(* IEC 61131-3 sources: IRIS-Project/LASAL CONTROL SOFTWARE/LasalProject_2025_09_12/Runtime/%LASALAPPDATA%/Runtime/Library/Loader/Source/code (part 10) *)

  OS_MT_Wait(pLogin^.hMutex);
  retval := SendLogout_TCP_nocs(pComdefT, pLogin);
  OS_MT_Signal(pLogin^.hMutex);

  UnlockLoginContext(pLogin); // wg. dem LockLoginContext2 Aufruf in dieser Funktion

END_FUNCTION
#endif

//------------------------------------------------------------------------------
// ComlinkT_InstallCallback
//------------------------------------------------------------------------------
#ifdef COMLINK_TCP_CLIENT
FUNCTION ComlinkT_InstallCallback
VAR_INPUT
    pCallback : ^void;
END_VAR
VAR
    i         : UDINT;
    pLogin    : ^loginContext;
END_VAR

  IF isClientReady < 0 THEN
    DEBUGLOG0("%010d-*** ComlinkT_InstallCallback: client is not ready");
    RETURN; // zeile geloescht laut pranz mail vom 30.01.2004
  END_IF;

  DEBUGLOG1("%010d-ComlinkT_InstallCallback: pCallback=0x%08X", pCallback$UDINT);

  FOR i := 0 TO (g_max_logins - 1) DO
    pLogin := LockLoginContext(i);
    IF pLogin <> NIL THEN
      pLogin^.pCallback := pCallback;
      UnlockLoginContext(pLogin);
    END_IF;
  END_FOR;

  g_pCallback := pCallback;

END_FUNCTION
#endif

//------------------------------------------------------------------------------
// ComlinkT_StartStopRefresh_nocs
//------------------------------------------------------------------------------
#ifdef COMLINK_TCP_CLIENT
FUNCTION ComlinkT_StartStopRefresh_nocs
VAR_INPUT
    pLogin   : ^loginContext; // connection context
    count    : UINT;
    typ      : UINT;
    res      : UDINT;
END_VAR
VAR_OUTPUT
    retval    : comlinkReason;
END_VAR
VAR
    reqMsg        : msgSsRefrReq;  // request structure for command CMD_SSREFR
    timeout_ms    : UDINT;         // timeout value for send request
    fFlush        : UDINT;
    rc            : DINT;
    rc2           : comlinkReason;
END_VAR

  retval := COMLINK_ERR_GENERAL;

  rc2 := CheckClientConnection(pLogin, #pLogin^.refrSockClnt, 0);
  IF rc2 <> COMLINK_OK THEN
    retval := rc2;
    RETURN;
  END_IF;

  // prepare the request message structure
  reqMsg.count   := count;
  reqMsg.typ     := typ;

  fFlush := 1;
  IF QUERY_FREE_TXBUF(pLogin^.refrSockClnt) < (2 * SIZEOF(reqMsg)) THEN
    DEBUGLOG0("%010d-*** ComlinkT_StartStopRefresh: send buffer shortage, next send will block");
    timeout_ms := CLIENT_TIMEOUT_REQ;
  ELSE
    timeout_ms := 0;    // timeout: non-blocking
  END_IF;

  pLogin^.accelerateCellUpdates := TRUE;

  // Send the request
  rc := SendCmdMsg(#pLogin^.refrSockClnt,
                   CMD_SSREFR,
                   0,                // Type and Ack field of command (type: request, ack: no response required)
                   #reqMsg$cMessage,
                   SIZEOF(reqMsg),
                   timeout_ms,
                   1,                // use buffered send
                   fFlush            // fFlush
                  );
  IF rc <= 0 THEN
    DEBUGLOG3("%010d-*** ComlinkT_StartStopRefresh(typ %d, count %d): SendCmdMsg failed, rc=%d", TO_UDINT(typ), TO_UDINT(count), TO_UDINT(rc));
    CloseBufferedSock(#pLogin^.refrSockClnt);
    retval := COMLINK_ERR_NOCONNECTION;
  ELSE
    DEBUG_VERBOSE3("%010d-ComlinkT_StartStopRefresh: SSREFR request sent, msgLen=%d, typ=%d, count=%d", TO_UDINT(rc), TO_UDINT(typ), TO_UDINT(count));
    retval := COMLINK_OK;
  END_IF;

END_FUNCTION
#endif

//------------------------------------------------------------------------------
// ComlinkT_StartStopRefresh
//------------------------------------------------------------------------------
#ifdef COMLINK_TCP_CLIENT
FUNCTION ComlinkT_StartStopRefresh
VAR_INPUT
    pComdef  : ^comdef;
    count    : UINT;
    typ      : UINT;
    res      : UDINT;
END_VAR
VAR_OUTPUT
    retval   : comlinkReason;
END_VAR
VAR
    pLogin        : ^loginContext; // connection context
END_VAR

  IF isClientReady < 0 THEN
    DEBUGLOG0("%010d-*** ComlinkT_StartStopRefresh: client is not ready");
    TraceMsg4Client();
    retval := COMLINK_ERR_CLIENT_NOTREADY;
    RETURN;
  END_IF;
  pLogin := pComdef^$comdefT.pLogin;
  IF pLogin = NIL THEN
    retval := COMLINK_ERR_LOGIN_REQUIRED;
    RETURN;
  END_IF;

  OS_MT_Wait(pLogin^.hMutex);
  retval := ComlinkT_StartStopRefresh_nocs(pLogin, count, typ, res);
  OS_MT_Signal(pLogin^.hMutex);

END_FUNCTION
#endif

//------------------------------------------------------------------------------
// ComlinkT_CyWork_Client - cyclic work for client
//------------------------------------------------------------------------------
#ifdef COMLINK_TCP_CLIENT
FUNCTION ComlinkT_CyWork_Client
VAR
    pLogin      : ^loginContext;
    reqMsgNop   : msgNopReq;
    rc          : DINT;
#ifndef LOADER_TCP_MODERATE
    i           : UDINT;
#endif
END_VAR

  IF (isClientReady < 0) | (loginAnz = 0) THEN
    RETURN;
  END_IF;

  TRACE_ENTRY(200);

#ifndef LOADER_TCP_MODERATE
  FOR i := 0 TO (g_max_logins - 1) DO

    pLogin := LockLoginContext(i);
#else
    pLogin := LockLoginContext(TCPCltCntr);
#endif

    IF pLogin <> NIL THEN

      TRACE_ENTRY(210);

      IF (pLogin^.cmdSockClnt.sock < 0) & (pLogin^.cmdSockClnt.pndSock >= 0) THEN
        // a pending command connection exists
        rc := Connect(pLogin^.cmdSockClnt.pndSock, pLogin^.ipAddrSrvr, pLogin^.cmdPortSrvr, 0);
        IF rc >= 0 THEN
          pLogin^.cmdSockClnt.sock    := pLogin^.cmdSockClnt.pndSock;
          pLogin^.cmdSockClnt.pndSock := INVALID_SOCKET_NUM;
          DEBUGLOG1("%010d-ComlinkT_CyWork: client connected to command server (port:%d)", pLogin^.cmdPortSrvr$UDINT);
        ELSIF rc <> TCP_NOT_READY THEN
          CloseSock(#pLogin^.cmdSockClnt.pndSock);
          DEBUGLOG2("%010d-ComlinkT_CyWork: connect to command server (port:%d) failed, rc=%d", pLogin^.cmdPortSrvr$UDINT, TO_UDINT(rc));
        END_IF;
      END_IF;

      IF (pLogin^.refrSockClnt.sock < 0) & (pLogin^.refrSockClnt.pndSock >= 0) THEN
        // a pending refresh connection exists
        rc := Connect(pLogin^.refrSockClnt.pndSock, pLogin^.ipAddrSrvr, pLogin^.cmdPortSrvr + 1, 0);
        IF rc >= 0 THEN
          pLogin^.refrSockClnt.sock    := pLogin^.refrSockClnt.pndSock;
          pLogin^.refrSockClnt.pndSock := INVALID_SOCKET_NUM;
          DEBUGLOG1("%010d-ComlinkT_CyWork: client connected to refresh server (port:%d)", (pLogin^.cmdPortSrvr + 1)$UDINT);
        ELSIF rc <> TCP_NOT_READY THEN
          CloseSock(#pLogin^.refrSockClnt.pndSock);
          DEBUGLOG2("%010d-ComlinkT_CyWork: connect to refresh server (port:%d) failed, rc=%d", (pLogin^.cmdPortSrvr + 1)$UDINT, TO_UDINT(rc));
        END_IF;
      END_IF;

      IF OS_MT_WaitCond(pLogin^.hMutex) THEN
        IF CheckClientConnection(pLogin, #pLogin^.refrSockClnt, 0) <> COMLINK_OK THEN

          TRACE_ENTRY(211);
          // poll for a response of the sessioninfo request
          PndConnListener(pLogin);

        ELSE

          TRACE_ENTRY(212);
          // flush the buffer when no transfer was in the last SMALLEST_UPD_INTERVALL ms
          IF (pLogin^.refrSockClnt.bytesInTxBuf > 0) &
             ((ops.tAbsolute - pLogin^.refrSockClnt.lastSendTime) > SMALLEST_UPD_INTERVALL) THEN
            DEBUG_VERBOSE1("%010d-ComlinkT_CyWork: initiate transfer of bufferd data (%d bytes)", pLogin^.refrSockClnt.bytesInTxBuf);
            FLUSH_TXBUF(#pLogin^.refrSockClnt);
          END_IF;

          // Send data at a regular interval to get informed when the server is not alive.
          // Without sending data at a regular interval we would recognize a connection failure
          // only when the LSE kernel initiates a transfer.
          // When we know that the server does not respond, we can initiate the reconnect procedure.
          IF (ops.tAbsolute - pLogin^.refrSockClnt.lastSendTime) > HEARTBEAT_INTERVALL THEN
            DEBUG_VERBOSE0("%010d-ComlinkT_CyWork: sending heartbeat");
            SendCmdMsg(#pLogin^.refrSockClnt, CMD_NOP, 0, #reqMsgNop$cMessage, SIZEOF(reqMsgNop), 0, 1, 1);
          END_IF;

          // send data in the buffer that is marked as unsent
          SendUnsentData(#pLogin^.refrSockClnt);

          // process incoming update cell requests
          IF ((ops.tAbsolute - pLogin^.refrSockClnt.lastUpdTime) > SMALLEST_UPD_INTERVALL) | pLogin^.accelerateCellUpdates THEN
            WHILE 1 DO
              IF UpdCellListener(pLogin) = 0 THEN
                // UpdCellListener returns 0 when no message is received
                EXIT;
              ELSE
                pLogin^.accelerateCellUpdates := FALSE;
              END_IF;
            END_WHILE;
            pLogin^.refrSockClnt.lastUpdTime := ops.tAbsolute;
          END_IF;

        END_IF;
        OS_MT_Signal(pLogin^.hMutex);
      END_IF; // OS_MT_WaitCond(pLogin^.hMutex)

      TRACE_ENTRY(219);

      UnlockLoginContext(pLogin);

    END_IF;

#ifdef LOADER_TCP_MODERATE
    TCPCltCntr += 1;
    if (TCPCltCntr = g_max_logins) then
      TCPCltCntr := 0;
    end_if;
#else
  END_FOR;
#endif

  TRACE_ENTRY(299);

END_FUNCTION
#endif

//------------------------------------------------------------------------------
// Ruft das Accept für den Command Socket auf
//------------------------------------------------------------------------------
#ifdef COMLINK_TCP_SERVER
FUNCTION ComlinkT_AcceptCmdSock
VAR
    sock        : DINT;
END_VAR

  IF cmdSockSrvr >= 0 THEN
    sock := OS_TCP_USER_ACCEPT(cmdSockSrvr, 0);
    IF sock >= 0 THEN
      DEBUGLOG1("%010d-  =====  command client connected  =====  , sock=%d", sock$UDINT);
      IF sock < arraysize(usedsocks) THEN
        usedsocks[sock] := 'C';
      END_IF;
      SetSocketOptions(sock);
      IF AllocConnBlock(TYPE_CMD_CONN, sock) = NIL THEN
        CloseSock(#sock);
      END_IF;
    END_IF;
  END_IF;

END_FUNCTION
#endif

//------------------------------------------------------------------------------
// Ruft das Accept für den Refresh Socket auf
//------------------------------------------------------------------------------
#ifdef COMLINK_TCP_SERVER
FUNCTION ComlinkT_AcceptRefrSock
VAR
    sock        : DINT;
END_VAR

  IF refrSockSrvr >= 0 THEN
    sock := OS_TCP_USER_ACCEPT(refrSockSrvr, 0);
    IF sock >= 0 THEN
      DEBUGLOG1("%010d-  =====  refresh client connected  =====  , sock=%d", sock$UDINT);
      IF sock < arraysize(usedsocks) THEN
        usedsocks[sock] := 'R';
      END_IF;
      SetSocketOptions(sock);
      IF AllocConnBlock(TYPE_REFR_CONN, sock) = NIL THEN
        CloseSock(#sock);
      END_IF;
    END_IF;
  END_IF;

END_FUNCTION
#endif

//------------------------------------------------------------------------------
// Serviciert einen offenen Command Socket
//------------------------------------------------------------------------------
#ifdef COMLINK_TCP_SERVER
FUNCTION ComlinkT_ServeCmdSock
VAR_INPUT
    pCmdConn    : ^cmdConnBlock;
END_VAR
#ifdef LOADER_TCP_MODERATE
VAR
	rc : DINT;
END_VAR
#endif

    // send data in the buffer that is marked as unsent
    SendUnsentData(#pCmdConn^.bsock);

    // process incoming command requests
    #ifdef LOADER_TCP_MODERATE
    rc :=
    #endif
    CmdMsgListener(pCmdConn);

    #ifdef LOADER_TCP_MODERATE
    IF rc >= 0 THEN
      pCmdConn^.bSock.isDataAvailable := false;
    END_IF;
    #endif

END_FUNCTION
#endif

//------------------------------------------------------------------------------
// Serviciert einen offenen Refresh Socket
//------------------------------------------------------------------------------
#ifdef COMLINK_TCP_SERVER
FUNCTION ComlinkT_ServeRefrSock
VAR_INPUT
    pRefrConn   : ^refrConnBlock;
END_VAR
VAR
    i           : UDINT;
    rc : DINT;
END_VAR

    // flush the buffer when no transfer was in the last SMALLEST_UPD_INTERVALL ms
    IF (pRefrConn^.bsock.bytesInTxBuf > 0) &
       ((ops.tAbsolute - pRefrConn^.bsock.lastSendTime) > SMALLEST_UPD_INTERVALL) THEN
      DEBUG_VERBOSE1("%010d-ComlinkT_CyWork: initiate transfer of bufferd data (%d bytes)", pRefrConn^.bsock.bytesInTxBuf);
      FLUSH_TXBUF(#pRefrConn^.bsock);
    END_IF;
    // send data in the buffer that is marked as unsent
    SendUnsentData(#pRefrConn^.bsock);

    // process incoming requests (TXUPD, StartStopRefresh)
    IF pRefrConn^.bsock.lastSendTime_ms <> ops.tAbsolute |
       pRefrConn^.bsock.refrMsgListenInhibitCnt > 5 // damit der RefrMsgListener auch eine Chance hat
       THEN
      // Es wird nur ein Receive durchgeführt, wenn in diesem Durchlauf nichts
      // gesendet wurde. Das begrenzt die CPU Last.
      i := 0;
      WHILE 1 DO
        rc := RefrMsgListener(pRefrConn);
        IF rc = 0 THEN
          // RefrMsgListener returns 0 when no message is received
          EXIT;
        END_IF;
        IF rc < 0 THEN
          // pRefrConn was released
          RETURN;
        END_IF;
        i += 1;
        IF i > 500 THEN // for safety
          EXIT;
        END_IF;
      END_WHILE;
      pRefrConn^.bsock.refrMsgListenInhibitCnt := 0;
    ELSE
      pRefrConn^.bsock.refrMsgListenInhibitCnt += 1;
    END_IF;
    // scan the update list and send changes to the client
    IF pRefrConn^.bsock.fTxBufferShortage THEN
      // no update in the case ot a buffer shortage
      IF QUERY_FREE_TXBUF(pRefrConn^.bsock) > (pRefrConn^.bsock.sizeOfTxBuf / 2) THEN
        DEBUGLOG0("%010d-ComlinkT_CyWork: leaving tx buffer shortage");
        pRefrConn^.bsock.fTxBufferShortage := 0;
      END_IF;
    ELSE
      IF ((ops.tAbsolute - pRefrConn^.bsock.lastUpdTime) > SMALLEST_UPD_INTERVALL) | pRefrConn^.flushNextSends THEN
        UpdateListProcessor(pRefrConn);
        pRefrConn^.bsock.lastUpdTime := ops.tAbsolute;
        IF pRefrConn^.flushNextSends THEN
          FLUSH_TXBUF(#pRefrConn^.bsock);
          pRefrConn^.flushNextSends := FALSE;
        END_IF;
      ELSE
        prefrconn := prefrconn;
      END_IF;
    END_IF;

    if( pRefrConn^.ptr = NIL )then
      return;
    end_if;
    IF pRefrConn^.ptr^.maxIdleTime_ms > 0 THEN
      IF ops.tAbsolute - pRefrConn^.bsock.lastSendTime_ms > pRefrConn^.ptr^.maxIdleTime_ms THEN
        SendAliveMessage_TCP(pRefrConn); // der Gegenstelle mitteilen, daß man noch lebt
      END_IF;
    END_IF;

END_FUNCTION
#endif

//------------------------------------------------------------------------------
// ComlinkT_CyWork_Server - cyclic work for server
//------------------------------------------------------------------------------
#ifdef COMLINK_TCP_SERVER
FUNCTION ComlinkT_CyWork_Server
VAR
    pCmdConnOld : ^cmdConnBlock;
    pRefrConnOld: ^refrConnBlock;
END_VAR

  IF isServerReady < 0 THEN
    RETURN;
  END_IF;

  // Die Aufrufe für das Accept des Kommando- und Refreshkanals und die
  // Bedienung dieser Kanäle wird so aufgeteilt, daß bei jedem Durchlauf
  // nur ein Aufruf gemacht wird, wobei die Accepts nur jedes 50te mal
  // aufgerufen werden. Ein Verbindungsaufbau braucht nämlich nicht so oft
  // überwacht werden.
  // Der Grund für diese Aufteilung ist der hohe CPU Verbrauch eines
  // TCP/IP Calls.

  CASE tcpServerState OF
    0:
      TRACE_ENTRY(100);
      // accept incoming command connection
      ComlinkT_AcceptCmdSock();
      tcpServerState += 1;

    1:
      TRACE_ENTRY(101);
      // accept incoming refresn connection
      ComlinkT_AcceptRefrSock();
      tcpServerState += 1;

    2:
      TRACE_ENTRY(102);
      // cyclic work for refresh server
      IF s_pRefrConn = NIL THEN
        s_pRefrConn := pRefrConnRoot;
      END_IF;
      IF s_pRefrConn <> NIL THEN

        ComlinkT_ServeRefrSock(s_pRefrConn);

        // check if an error occured
        IF s_pRefrConn <> NIL THEN // s_pRefrConn kann in ComlinkT_ServeRefrSock freigegeben werden
	        IF s_pRefrConn^.bsock.sock < 0 THEN
	          pRefrConnOld := s_pRefrConn;
	          s_pRefrConn    := s_pRefrConn^.next;
            DEBUGLOG0("%010d-  =====  Error in RefrConn -> releasing connBlock  =====");
	          ReleaseConnBlock(TYPE_REFR_CONN, pRefrConnOld$^connBlock, 1);
            pRefrConnOld := NIL;
	        ELSE
	          s_pRefrConn := s_pRefrConn^.next;
	        END_IF;
        END_IF;

      END_IF;
      IF s_pRefrConn = NIL THEN
        tcpServerState += 1;
      END_IF;

    3:
      TRACE_ENTRY(103);
      // cyclic work for command server
      IF s_pCmdConn = NIL THEN
        s_pCmdConn := pCmdConnRoot;
      END_IF;
      IF s_pCmdConn <> NIL THEN

        ComlinkT_ServeCmdSock(s_pCmdConn);

        // check if an error occured
        IF s_pCmdConn <> NIL THEN // s_pCmdConn kann in ComlinkT_ServeCmdSock freigegeben werden
	        IF s_pCmdConn^.bsock.sock < 0 THEN
	          pCmdConnOld := s_pCmdConn;
	          s_pCmdConn    := s_pCmdConn^.next;
            DEBUGLOG0("%010d-  =====  Error in CmdConn -> releasing connBlock =====");
	          ReleaseConnBlock(TYPE_CMD_CONN, pCmdConnOld$^connBlock, 0);
            pCmdConnOld := NIL;
	        ELSE
	          s_pCmdConn := s_pCmdConn^.next;
	        END_IF;
        END_IF;

      END_IF;
      IF s_pCmdConn = NIL THEN
        tcpServerState += 1;
      END_IF;

  END_CASE;

  tcpAcceptState += 1;

  IF tcpServerState > 3 THEN
    // Es wird nur alle 50 Durchläufe ein Accept eingeschoben
    IF tcpAcceptState > 50 THEN
      tcpAcceptState := 0;
      tcpServerState := 0;
    ELSE
      tcpServerState := 2;
    END_IF;
  END_IF;

  TRACE_ENTRY(199);

END_FUNCTION
#endif

//------------------------------------------------------------------------------
// ComlinkT_CyWork
//------------------------------------------------------------------------------
FUNCTION ComlinkT_CyWork

  TRACE_ENTRY(10);

#ifdef COMLINK_TCP_SERVER
  ComlinkT_CyWork_Server();
#endif

  TRACE_ENTRY(11);

#ifdef COMLINK_TCP_CLIENT
  ComlinkT_CyWork_Client();
#endif

  TRACE_ENTRY(12);

END_FUNCTION

#endif //COMLINK_TCP

#ifndef COMLINK_TCP_CLIENT

//------------------------------------------------------------------------------
// ComlinkT_MissingClientCode
//------------------------------------------------------------------------------
FUNCTION ComlinkT_MissingClientCode

  IF ComlinkT_wasTraceMsgDisplayed = 0 THEN
    TRACE_ERR("Comlink/TCP client error: missing client code (COMLINK_TCP_CLIENT not defined)");
    LSLCLI_LoaderTracePrint("Comlink/TCP client error: missing client code (COMLINK_TCP_CLIENT not defined)", 12);
    ComlinkT_wasTraceMsgDisplayed := 1;
  END_IF;

END_FUNCTION

#endif // !COMLINK_TCP_CLIENT

//++comlinkt:end

////////////////////////////////////////////////////////////////////////////////
//
//  I-am-Alive Mechanismus
//
////////////////////////////////////////////////////////////////////////////////

FUNCTION SendMaxIdleTime_CAN
VAR_INPUT
  pComdefT : ^comdefT;
  remoteMaxIdleTime_ms : UDINT;
END_VAR
VAR_OUTPUT
  retVal : DINT;
END_VAR
VAR
  txinfo4006    : COMOBJSTR;
END_VAR

    txinfo4006.iLng  := 0;
    txinfo4006.iOff  := 4006;
    txinfo4006.dData := TO_DINT(remoteMaxIdleTime_ms);

    IF CanTxObj(pComdefT$^COMDEF^.pt_COM, #txinfo4006$void) <> 0 THEN
        retVal := -1;
    ELSE
        retVal := 0;
    END_IF;

END_FUNCTION
FUNCTION SendAliveMessage_CAN
VAR_INPUT
  pCom : ^COMDATA;
END_VAR
VAR_OUTPUT
  retVal : DINT;
END_VAR
VAR
  txinfo4007    : COMOBJSTR;
END_VAR

    txinfo4007.iLng  := 0;
    txinfo4007.iOff  := 4007;
    txinfo4007.dData := 0;

    IF CanTxObj(pCom, #txinfo4007$void) <> 0 THEN
        retVal := -1;
    ELSE
        retVal := 0;
    END_IF;

END_FUNCTION
//------------------------------------------------------------------------------
// SendMaxIdleTime
//
//  Schickt die maxIdleTime zur Gegenstation
//------------------------------------------------------------------------------
FUNCTION SendMaxIdleTime
VAR_INPUT
  pComdefT : ^comdefT;
  remoteMaxIdleTime_ms : UDINT;
END_VAR
VAR_OUTPUT
  retVal : DINT;
END_VAR

  CASE pComdefT^.interface  OF

  COMLINK_IFNUM_CAN1,
  COMLINK_IFNUM_CAN2,
  COMLINK_IFNUM_CAN20,
  COMLINK_IFNUM_CAN21,
  COMLINK_IFNUM_CAN22,
  COMLINK_IFNUM_CAN23,
  COMLINK_IFNUM_CAN24,
  COMLINK_IFNUM_CAN25,
  COMLINK_IFNUM_CAN26,
  COMLINK_IFNUM_CAN27,
  COMLINK_IFNUM_CAN28,
  COMLINK_IFNUM_CAN29:
    retVal := SendMaxIdleTime_CAN(pComdefT, remoteMaxIdleTime_ms);
#ifdef COMLINK_TCP_SERVER
  COMLINK_IFNUM_TCP1_OLD,
  COMLINK_IFNUM_TCP1,
  COMLINK_IFNUM_TCP2:
    retVal := SendMaxIdleTime_TCP(pComdefT, remoteMaxIdleTime_ms);
#endif
  COMLINK_IFNUM_COM1,
  COMLINK_IFNUM_COM2,
  COMLINK_IFNUM_COM3,
  COMLINK_IFNUM_COM4,
  COMLINK_IFNUM_COM5,
  COMLINK_IFNUM_COM6,
  COMLINK_IFNUM_COM7,
  COMLINK_IFNUM_COM8,
  COMLINK_IFNUM_COM9,
  COMLINK_IFNUM_COM10:
    retVal := SendMaxIdleTime_RS232(pComdefT, remoteMaxIdleTime_ms);
  ELSE
    retVal := -1;
  END_CASE;

END_FUNCTION

//------------------------------------------------------------------------------
// SendMaxIdleTime
//
//  Schickt die maxIdleTime zur Gegenstation
//------------------------------------------------------------------------------
FUNCTION SendLogout
VAR_INPUT
  pComdefT : ^comdefT;
END_VAR
VAR_OUTPUT
  retVal : DINT;
END_VAR

  CASE pComdefT^.interface  OF

  COMLINK_IFNUM_CAN1,
  COMLINK_IFNUM_CAN2,
  COMLINK_IFNUM_CAN20,
  COMLINK_IFNUM_CAN21,
  COMLINK_IFNUM_CAN22,
  COMLINK_IFNUM_CAN23,
  COMLINK_IFNUM_CAN24,
  COMLINK_IFNUM_CAN25,
  COMLINK_IFNUM_CAN26,
  COMLINK_IFNUM_CAN27,
  COMLINK_IFNUM_CAN28,
  COMLINK_IFNUM_CAN29:
    //retVal := SendMaxIdleTime_CAN(pComdefT, remoteMaxIdleTime_ms);
#ifdef COMLINK_TCP_SERVER
  COMLINK_IFNUM_TCP1_OLD,
  COMLINK_IFNUM_TCP1,
  COMLINK_IFNUM_TCP2:
    retVal := SendLogout_TCP(pComdefT);
#endif
  COMLINK_IFNUM_COM1,
  COMLINK_IFNUM_COM2,
  COMLINK_IFNUM_COM3,
  COMLINK_IFNUM_COM4,
  COMLINK_IFNUM_COM5,
  COMLINK_IFNUM_COM6,
  COMLINK_IFNUM_COM7,
  COMLINK_IFNUM_COM8,
  COMLINK_IFNUM_COM9,
  COMLINK_IFNUM_COM10:
    //retVal := SendMaxIdleTime_RS232(pComdefT, remoteMaxIdleTime_ms);
  ELSE
    retVal := -1;
  END_CASE;

END_FUNCTION

//------------------------------------------------------------------------------
// AliveCheck
//
//  Überprüft bei einem Node:
//  a) ob die Zeit maxSilentTime_ms abgelaufen ist (dann wird angenommen, daß
//     die Gegenstelle tot ist oder die Verbindung unterbrochen wurde)
//  b) ob der Gegenstelle eine Alive-Message geschickt worden ist (falls seit
//     der letzten gesendeten Message schon zu viel Zeit vergangen ist)
//------------------------------------------------------------------------------
FUNCTION AliveCheck
VAR_INPUT
    pNode : ^MonitorNode;
END_VAR

    IF pNode^.maxSilentTime_ms > 0 THEN
        IF ops.tAbsolute - pNode^.lastRcvdTime_ms > pNode^.maxSilentTime_ms THEN
            pNode^.isRemotePlcAlive := FALSE;   // Flag, das anzeigt, daß die Gegenstelle nicht mehr antwortet
        END_IF;
    END_IF;

END_FUNCTION

//------------------------------------------------------------------------------
// AliveChecker
//
//  Geht die Liste aller zu überwachenden Nodes durch und ruft für jeden Node
//  die Funktion AliveCheck auf.
//------------------------------------------------------------------------------
FUNCTION AliveChecker
VAR
  pWork : ^MonitorNodeList;
END_VAR

  // die folgende Abfrage vermeidet die Verwendung des monitorNodeMutex wenn nichts
  // zu überwachen ist
  IF monitorNodes = NIL THEN
    RETURN;
  END_IF;

  OS_MT_WAIT(monitorNodeMutex);

  pWork := monitorNodes;
  WHILE pWork DO
    AliveCheck(pWork$^MonitorNode);
    pWork := pWork^.pNext;
  END_WHILE;

  OS_MT_SIGNAL(monitorNodeMutex);

END_FUNCTION
//------------------------------------------------------------------------------
// SearchMonitorNode
//
//  Sucht einen Node in der Überwachungsliste anhand der in pComdefT
//  gespeicherten Netzwerkadresse .
//------------------------------------------------------------------------------
(*

    Diese Funktion kann man verwenden, wenn man nicht pro Kanal sondern pro
    Netzwerkadresse überwacht.

FUNCTION SearchMonitorNode
VAR_INPUT
  pComdefT : ^comdefT;
END_VAR
VAR_OUTPUT
  pNode : ^MonitorNode;
END_VAR
VAR
  pWork : ^MonitorNodeList;
END_VAR

  pNode := NIL;
  pWork := monitorNodes;

  WHILE pWork DO

    CASE pComdefT^.interface  OF

    COMLINK_IFNUM_CAN1:
      IF pComdefT^.canAddress = pWork$^MonitorNode^.canAddress THEN
        pNode := pWork$^MonitorNode;
        EXIT;
      END_IF;

    COMLINK_IFNUM_TCP1_OLD,
    COMLINK_IFNUM_TCP1,
    COMLINK_IFNUM_TCP2:
      IF pComdefT^.ipAddress = pWork$^MonitorNode^.ipAddress &
         pComdefT^.port      = pWork$^MonitorNode^.port THEN
        pNode := pWork$^MonitorNode;
        EXIT;
      END_IF;
    END_CASE;

    pWork := pWork^.pNext;
  END_WHILE;

END_FUNCTION
*)

//------------------------------------------------------------------------------
// RemoveMonitorNode
//
//  Hängt einen Node aus der Überwachungsliste aus
//------------------------------------------------------------------------------
FUNCTION RemoveMonitorNode
VAR_INPUT
  pNode : ^MonitorNode;
END_VAR
VAR
  pPrev : ^MonitorNodeList;
  pWork : ^MonitorNodeList;
END_VAR

  pPrev := NIL;
  pWork := monitorNodes;

  WHILE pWork DO

    IF pWork$^MonitorNode = pNode THEN
      IF pPrev = NIL THEN
        monitorNodes := pWork^.pNext;
      ELSE
        pPrev^.pNext := pWork^.pNext;
      END_IF;
      _free(pWork);
      pWork := NIL;
      EXIT;
    END_IF;

    pPrev := pWork;
    pWork := pWork^.pNext;
  END_WHILE;

END_FUNCTION

//------------------------------------------------------------------------------
// AddMonitorNode
//
//  Hängt einen Node in die Überwachungsliste ein
//------------------------------------------------------------------------------
FUNCTION AddMonitorNode
VAR_INPUT
    pNode : ^MonitorNode;
END_VAR

    pNode$^MonitorNodeList^.pNext := monitorNodes;
    monitorNodes := pNode$^MonitorNodeList;

END_FUNCTION
//------------------------------------------------------------------------------
// DeactivateAliveCheck
//
//  Deaktiviert die Überwachung einer Comlink Gegenstelle.
//------------------------------------------------------------------------------
FUNCTION DeactivateAliveCheck
VAR_INPUT
  pComdefT : ^comdefT;
END_VAR
VAR_OUTPUT
  retVal : DINT;
END_VAR
VAR
  pt_COM   : ^COMDATA;
  pNode : ^MonitorNode;
END_VAR

  retVal := SendMaxIdleTime(pComdefT, 0);

  pt_COM := pComdefT^.pLogin$^COMDATA;
  IF pt_COM <> NIL THEN
    OS_MT_WAIT(monitorNodeMutex);
    IF pt_COM^.pNode THEN
      pNode := pt_COM^.pNode;
      pt_COM^.pNode := NIL;
      RemoveMonitorNode(pNode);
    END_IF;
    OS_MT_SIGNAL(monitorNodeMutex);
  END_IF;

END_FUNCTION
//------------------------------------------------------------------------------
// ActivateAliveCheck
//
//  Aktiviert die Überwachung einer Comlink Gegenstelle. Der Timeout für die
//  Überwachung wird mit dem Parameter maxSilentTime_ms angegeben.
//  remoteMaxIdleTime_ms wird der Gegenstelle mitgeteilt.
//------------------------------------------------------------------------------
FUNCTION ActivateAliveCheck
VAR_INPUT
  pComdefT : ^comdefT;
  maxSilentTime_ms : UDINT;
  remoteMaxIdleTime_ms : UDINT;
END_VAR
VAR_OUTPUT
  retVal : DINT;
END_VAR
VAR
    pt_COM   : ^COMDATA;
    pNode : ^MonitorNode;
    pOldNode : ^MonitorNode;
END_VAR

    retVal := 0;

    pt_COM := pComdefT^.pLogin$^COMDATA;
    IF pt_COM = NIL THEN
      RETURN;
    END_IF;

    OS_MT_WAIT(monitorNodeMutex);
    pOldNode := pt_COM^.pNode;
    IF pOldNode = NIL THEN
        // für diesen Kanal war noch kein Eintrag vorhanden -> neuen Listeneintrag erstellen
        pNode := calloc(SIZEOF(MonitorNodeList))$^MonitorNode;
        IF pNode <> NIL THEN
            pNode^.pt_COM           := pt_COM;
            pNode^.isRemotePlcAlive := TRUE;
        END_IF;
    ELSE
        // bestehenden Listeneintrag wiederverwenden
        pNode := pOldNode;
    END_IF;
    OS_MT_SIGNAL(monitorNodeMutex);

    IF pNode = NIL THEN
        retVal := -1;
        RETURN;
    END_IF;

    (*
    // prüfen, ob die bisherigen Einstellungen des Nodes geändert werden müssen
    -> nur notwendig, wenn pro Netzwerkadresse und nicht pro Kanal überwacht wird
    IF pOldNode = NIL | maxSilentTime_ms < pNode^.maxSilentTime_ms THEN
        IF pOldNode = NIL | remoteMaxIdleTime_ms <> pNode^.remoteMaxIdleTime_ms THEN
            // Es wurde entweder ein neuer Eintrag in der Überwachungsliste erstellt
            // oder der neue Wert für die maxIdleTime ist anders als der bisherige.
            pNode^.remoteMaxIdleTime_ms := remoteMaxIdleTime_ms;
        END_IF;
        pNode^.maxSilentTime_ms := maxSilentTime_ms;
    END_IF;
    *)

    // Der neue Wert für remoteMaxIdleTime_ms wird in jedem Fall gesendet, auch
    // wenn man annehmen müßte daß die Gegenstelle den aktuellen Wert schon hat.
    // Wenn nämlich die Gegenstelle resettiert worden ist, dann hat sie die Einstellungen
    // vergessen.
    retVal := SendMaxIdleTime(pComdefT, remoteMaxIdleTime_ms);
    IF retVal < 0 THEN
        IF pOldNode = NIL THEN
            _free(pNode);
            pNode := NIL;
            RETURN;
        END_IF;
    END_IF;

    OS_MT_WAIT(monitorNodeMutex);
    pNode^.lastRcvdTime_ms := ops.tAbsolute;
    pNode^.maxSilentTime_ms := maxSilentTime_ms;
    pNode^.remoteMaxIdleTime_ms := remoteMaxIdleTime_ms;

    IF pOldNode = NIL THEN
        // neuen Node in die Überwachungs-Liste einhängen
        AddMonitorNode(pNode);
    END_IF;

    // Die Zeit-Werte merken, damit beim entfernen eines Nodes aus der Überwachungs-Liste
    // ein passender neuer Eintrag gesucht werden kann.
    pt_COM^.pNode := pNode;
    OS_MT_SIGNAL(monitorNodeMutex);

END_FUNCTION
//------------------------------------------------------------------------------
// LDR_SetIamAliveTime
//
//  API Funktion zum aktivieren oder deaktivieren der Überwachung einer Comlink
//  Gegenstelle.
//
//  pComdefT
//    Comdef Struktur der Comlink Verbindung
//  remoteMaxIdleTime_ms
//    'maxIdleTime' die der Gegenstelle mitgeteilt wird. Die Gegenstelle schickt
//    eine Message, wenn sie feststellt daß seit der letzten gesendeten Message
//    die Zeit 'maxIdleTime' vergangen ist.
//      >0  .. Wert in ms
//      -1  .. Default-Wert (100ms),
//       0  .. deaktivieren
//  maxNetworkDelay_ms
//    Die maximale Netzwerkverzögerung für diese Verbindung.
//     >=0  .. Wert in ms
//      -1  .. Default-Wert (20ms),
//  remoteMaxCyclicTime_ms
//    Die max.Durchlaufzeit des Cyclics der Gegenstation (nur für den Fall daß
//    die Gegenstelle diesen Wert nicht liefert).
//     >=0  .. Wert in ms
//      -1  .. Default-Wert (300ms),
//
//  Return:
//    0  .. o.k.
//   <0  .. Fehler
//------------------------------------------------------------------------------
FUNCTION GLOBAL __CDECL LDR_SetIamAliveTime
VAR_INPUT
  pComdef : ^COMDEF;
  remoteMaxIdleTime_ms : UDINT;
  maxNetworkDelay_ms : UDINT;
  remoteMaxCyclicTime_ms : UDINT;
END_VAR
VAR_OUTPUT
  retVal : DINT;
END_VAR

    IF (pComdef = NIL) | (pComdef^.pt_Com = NIL) THEN
        retVal := -1;
        RETURN;
    END_IF;

    IF pComdef^.pt_COM^.remoteMaxCyclicTime_ms = 16#FFFFffff THEN
        // die Gegenstelle hat beim Login keine maxCyclicTime geschickt,
        // d.h. daß die Loaderversion der Gegenstelle den Alive Mechanismus
        // noch nicht implementiert hat. -> Fehlercode zurückgeben
        retVal := -1;
        RETURN;
    END_IF;

    IF remoteMaxIdleTime_ms = 0 THEN
        // Überwachung deaktivieren
        retVal := DeactivateAliveCheck(pComdef$^comdefT);
    ELSE
        // Defaultwerte übernehmen
        IF remoteMaxIdleTime_ms = 16#FFFFffff THEN
            remoteMaxIdleTime_ms := 100;
        END_IF;
        IF maxNetworkDelay_ms = 16#FFFFffff THEN
            maxNetworkDelay_ms := 20;
        END_IF;
        IF pComdef^.pt_COM^.remoteMaxCyclicTime_ms <> 0 THEN
            // die Gegenstelle hat für ihre eigene maxCyclicTime einen Wert <> 0 mitgeteilt
            remoteMaxCyclicTime_ms := pComdef^.pt_COM^.remoteMaxCyclicTime_ms;
        ELSIF remoteMaxCyclicTime_ms = 16#FFFFffff THEN
            // maxCyclicTime ist weder vom Aufrufer noch von der Gegenstelle mitgeteilt worden
            // -> Defaultwert verwenden.
            remoteMaxCyclicTime_ms := 300;
        END_IF;

        // Überwachung aktivieren
        retVal := ActivateAliveCheck(pComdef$^comdefT,
                                     remoteMaxIdleTime_ms + maxNetworkDelay_ms + remoteMaxCyclicTime_ms,
                                     remoteMaxIdleTime_ms);
    END_IF;

END_FUNCTION
//------------------------------------------------------------------------------
// LDR_isRemotePlcAlive
//
//  Mit dieser API Funktion kann festgestellt werden, ob von der Remote PLC
//  regelmäßig etwas geschickt wird.
//
//  Return:
//    0  .. Die Remote PLC hat sich in letzter Zeit nicht mehr gemeldet
//   >0  .. Von der Remote PLC werden regelmäßig Daten empfangen
//------------------------------------------------------------------------------
FUNCTION GLOBAL __CDECL LDR_isRemotePlcAlive
VAR_INPUT
  pComdef : ^COMDEF;
END_VAR
VAR_OUTPUT
  retVal : DINT;
END_VAR

    retVal := 0;
    IF pComdef & pComdef^.pt_COM & pComdef^.pt_COM^.pNode  THEN
        retVal := pComdef^.pt_COM^.pNode^.isRemotePlcAlive;
    END_IF;

END_FUNCTION
//------------------------------------------------------------------------------
// LDR_SetCanWait
//------------------------------------------------------------------------------
FUNCTION GLOBAL __CDECL LDR_SetCanWait //ws001
VAR_INPUT
  us_wait : usint;
END_VAR
VAR_OUTPUT
  old : usint;
END_VAR

  old := LDR_canwait;
  LDR_canwait := us_wait;

END_FUNCTION // /ws001
//------------------------------------------------------------------------------
// LDR_SetWait4Visu
//  Setzt das Flag bWait4Visu. Wenn dieses Flag gesetzt ist, dann wird nach der
//  Loader-Initialisierung nicht sofort der zyklische Betrieb aufgenommen.
//  Dadurch bleibt mehr CPU Zeit für die GetId-Phase der Visu übrig und die
//  GetId-Phase wird schneller fertig.
//  Der zyklische Betrieb wird dann gestartet, wenn das Flag bWait4Visu (siehe
//  Befehl I_VISU_RDY) wieder zurückgesetzt wird. Mit dem Parameter timeout_ms
//  kann ein Timeout-Wert festgelegt werden, nach dem der zyklische Betrieb
//  aufgenommen wird, auch wenn das Flag bWait4Visu nicht zurückgesetzt wird.
//  Der Timeout-Wert 0 bedeutet dass der Timeout nicht wirksam ist.
//------------------------------------------------------------------------------
FUNCTION GLOBAL __CDECL LDR_SetWait4Visu  //ZP000
VAR_INPUT
  bWait : BOOL;
  timeout_ms : UDINT;
END_VAR

  bWait4Visu := bWait;
  wait4Visu_timeout_ms := timeout_ms;

END_FUNCTION  //ZP000
//------------------------------------------------------------------------------
// LDR_SetCanWaitRemote
//
//  Legt den Wert der Canbremse serverseitig fest (nur für diesen einen Kanal).
//  -1 bedeutet Defaultwert wiederherstellen.
//------------------------------------------------------------------------------
FUNCTION GLOBAL __CDECL LDR_SetCanWaitRemote
VAR_INPUT
  pComdef : ^COMDEF;
  wait : INT;
END_VAR
VAR_OUTPUT
  retVal : DINT;
END_VAR
VAR
  txinfo4008    : COMOBJSTR;
END_VAR

    txinfo4008.iLng  := 0;
    txinfo4008.iOff  := 4008;
    txinfo4008.dData := 0;
    txinfo4008.dData$INT := wait;

    IF CanTxObj(pComdef^.pt_COM, #txinfo4008$void) <> 0 THEN
        retVal := -1;
    ELSE
        retVal := 0;
    END_IF;

END_FUNCTION

(*===============================================================================

  ComlinkRS232 - Comlink über RS232

===============================================================================*)

(*
  Konzept:
  --------

  Auf unterer Ebene (L0) werden L0-Pakete (L0-Requests und L0-Responses) hin- und
  hergeschickt. Der Aufbau ist so gewählt, daß sich die L0-Pakete mit dem Lasal32
  Protokoll vertragen, d.h. wenn das Lasal32 Protokoll Comlink Daten empfängt
  (oder umgekehrt), dann wird das Paktetformat verstanden, das darin enthaltene
  Kommandobyte wird aber als nicht unterstützter Befehl erkannt und es wird ein
  NAK zurückgeschickt.

  In einem L0-Paket sind die Comlink Requests und Responses eingepackt (z.B.
  TxCommand Req.+Resp., UpdCell Req. usw.).

  Ein L0-Paket ist mit einer Checksumme versehen, um Übertragungsfehler zu
  erkennen.

  Wenn ein L0-Request geschickt wird, dann muss auf die L0-Response gewartet werden,
  bis wieder ein L0-Request geschickt werden darf. Wenn ein L0-Request empfangen
  wird, dann muss dieser mit einer L0-Response beantwortet werden, sonst schickt
  die Gegenstation nichts mehr. Mit diesem Mechanismus erreicht man eine Fluss-
  kontrolle, d.h. man kann den Empfangsbuffer der Gegenstation nicht überfluten.
  Der Empfangsbuffer der Gegenstation muss so gross gewählt werden, daß er mindestens
  den größtmöglichen L0-Request und die größtmöglichen L0-Response aufnehmen kann.
  Die Werte wurden so gewählt, daß ein L0-Paket (Req. oder Resp.) max. 1000 Bytes
  gross sein kann, daher muss der Empfangsbuffer 2000 Bytes gross sein.

  Die Comlink Requests und Responses sind L1 Pakete. Es gibt L0-Sendebuffer,
  in welche die zu sendenden L1 Pakete beim Sendeaufruf hineingestellt werden.
  In einen L0-Sendebuffer können nur dann L1 Pakete hineinkopiert werden, wenn
  er nicht gerade vom Sendeteil in Bearbeitung ist.
  Es werden 2 L0-Sendebuffer verwendet, damit auch Daten entgegengenommen werden
  können, wenn einer in Bearbeitung ist (solange bis dieser freie L0-Sendebuffer
  voll ist).

  Thread-Sicherheit:
  - Funktionsaufrufe für verschiedene Kanäle können aus verschiedenenen Tasks
    aufgerufen werden.
  - Bei Funktionsaufrufen für den gleichen Kanal können nur Befehle aus unterschiedlichen
    Befehlsgruppen aus verschiedenen Tasks aufgerufen werden.
    Es gibt 2 Befehlsgruppen: Command- und Refreshlistenbefehle.
    Commandbefehl: TxCommand
    Refreshbefehl: TxUpd, StartStopRefresh
*)

#define NBR_OF_RS232_ITFS 10   // Anzahl der unterstützten RS232 Schnittstellen

#define DFLT_BAUD         9
#define DFLT_PARITY       0
#define DFLT_STOP         1
#define DFLT_WORDL        8

TYPE

#pragma pack (push,1)

#define L0_STX   16#02
#define L0_ETX   16#03

#define RS232_L0_TIMEOUT_BAUD115KB          500  // bezogen auf 115200 baud (in dieser Zeit können ca. 5 1k Pakete übertragen werden)
#define RS232_L0_TIMEOUT_GSMDELAY          1000  // Verzögerung wenn ein GSM Modem verwendet wird

#define RS232_L0_RESP_TIMEVAL               100  // nach dieser Zeit wird spätestens eine L0 Response geschickt

#define RS232_L0FLAGS_IS_REQUEST          16#01
#define RS232_L0CMD                       16#A0

#define L0_EMPTY_DATALEN    5   // Das ist die DataLen im L0 Header, wenn 0 Bytes Schicht1 Daten vorhanden sind (nur HdrChk ist vorhanden)

  // Schicht 0 Datenformat
  // !STX  !                       !0xA0 !Hdr  !<---  Schicht1 Daten  --->!  Data     !ETX  !
  // !0x02 !        DataLen        !Flags!Chk  !            ...           !  Chksum   !0x03 !
  // +-----+-----+-----+-----+-----+-----+-----+-----+-----         +-----+-----+-----+-----+
  //        \-------- Hdr Chksum -------/ \--------  DataLen-4  ---------/
  //                                \----------- Data Chksum ------------/
  //  \------------------------------- DataLen+5 ------------------------------------------/
  SER_L0_BUF : STRUCT
    stx : BYTE;
    dataLen : UDINT;
    flagsCmd : BYTE;
    hdrChksum : BYTE;
    data : ARRAY[0..992] OF BYTE; // Platz für 990 Datenbytes, 2 Bytes Chksum, 1 Byte ETX
  END_STRUCT;

#define INVALID_CHIDX   254
#define UNKNOWN_CHIDX   255

#define RS232_L1CMD_MASK    16#3F

#define RS232_L1FLAGS_IS_REQUEST          16#80
#define RS232_L1FLAGS_RESPONSE_REQUIRED   16#40 // nur bei einem Request relevant
#define RS232_L1FLAGS_ACK                 16#40 // nur bei einer Response relevent (0=unbekannter Befehl)
  // Schicht 1 Datenformat
  // !Src  !Dst  !Flags!           !           !                             !
  // !ChIdx!ChIdx!Cmd  !  DataLen  !  Seq.Nbr  !  Data       ...             !
  // +-----+-----+-----+-----+-----+-----+-----+-----+-----+     +-----+-----+
  //                                \--------------- DataLen ---------------/
  SER_L1_TXBUF : STRUCT
    dataValid : BYTE; // wird nicht gesendet !
    srcChIdx : BYTE;
    dstChIdx : BYTE;
    flagsCmd : BYTE;
    dataLen : UINT;
    data : ARRAY[0..299] OF BYTE;
  END_STRUCT;

  SER_L1_BUF : STRUCT
    srcChIdx : BYTE;
    dstChIdx : BYTE;
    flagsCmd : BYTE;
    dataLen : UINT;
    data : ARRAY[0..299] OF BYTE;
  END_STRUCT;
#pragma pack (pop)

  RS232_ITF : STRUCT
    hComm : pVoid;              // Handle für die RS232 Schnittstelle
    hCommAppl : pVoid;          // das gleiche Handle - wird während der Initialisierungsphase von der Applikation verwendet (z.B.Modem Wählvorgang)
    baudrate : UINT;            // zu verwendende Baudrate
    timeoutVal : UDINT;         // Timeout in ms
    startServer : DINT;         // Flag, ob der Comlink Server die Schnittstelle benutzen soll
    fnInitInterface : pVoid;    // Callbackfunktion in der z.B. einen Modemverbindung aufgebaut wird
    pThis : pVoid;              // This-Pointer für die Callbackfunktion

    itfIdx : DINT;              // Index im rs232Itfs Array

    l0SendBufA : SER_L0_BUF;
    l0SendBufB : SER_L0_BUF;

    pL0SendBufferCollect : ^SER_L0_BUF;
    pL0SendBufferTransfer : ^SER_L0_BUF;
    bytesToSend : UDINT;        // Anzahl der zu sendenden Bytes im pL0SendBufferTransfer
    bytesSent : UDINT;          // Anzahl der gesendeten Bytes im pL0SendBufferTransfer
    sendInProgress : BOOL;      // TRUE, wenn das Senden läuft

    l0RespPending : BOOL;       // es wird eine L0 Response erwartet
    l0RespNecessary : BOOL;     // es muss eine L0 Response geschickt werden
    l0RespPendingTimeout_ms : UDINT;    // Wenn nach dieser Zeit keine Resp. eintrifft, dann wird das Flag zurückgesetzt
    l0RespNecessaryTimeval_ms : UDINT;  // Wenn nach dieser Zeit noch keine Resp. geschickt wurde, dann wird eine Response auch ohne Daten geschickt

    bytesInRecvBuf : UDINT;
    l0RecvBuf : ARRAY[0..999] OF BYTE;  // L0-Empfangsbuffer
  END_STRUCT;

#pragma pack (push,1)
  loginContextR : STRUCT
    // ---- muß immer da vorne sein (wegen CAN comData Structur) ----
    pCallback                     : ^void;
    pThis                         : UDINT;
    hComchMutex                   : MT_SEMAHANDLE; //
    typeOfStruct				          : UINT;		   // STRUCT_TYPE_...
    sizeofDynList                 : UINT;          //
    sizeofStatList                : UINT;          //
    sizeofRemoteDynList           : UINT;          //
    sizeofRemoteStatList          : UINT;          //
    remoteMaxCyclicTime_ms        : UDINT;         //
    pNode                         : ^MonitorNode;  //
    pDynCallbacks       		  : ^sDynCallbackList; // Liste der Callbacks (ua. für Multimaster)
    // ---------------------------------------------------------
    versionOfPeer: UDINT;           // version number of the peer
    instIdOfPeer : UDINT;           // instance id of the peer
    interface    : UDINT;           // interface nummer (kein Index, nicht 0-basierend !)
    pItf         : ^RS232_ITF;

    txL1BufCmd   : SER_L1_TXBUF;    // der Sendebuffer für TxCommand, bzw. die Response darauf
    txL1BufRefr  : SER_L1_TXBUF;    // der Sendebuffer für die Verwaltung der Updatelisten
    rxL1BufResp  : SER_L1_BUF;
    rxL1BufReq   : SER_L1_BUF;
    statList     : updateList;      // static list
    dynList      : updateList;      // dynamic list
    pComdefT     : ^comdefT;        // a pointer to a structure that was given by the caller of login
    hMutex       : MT_SEMAHANDLE;   // Mutex for ???
    myChIdx      : BYTE;            // Channel Index lokal
    hisChIdx     : BYTE;            // Channel Index remote
    isConnected  : BOOL;            // nach einem Login:connected, nach einem Fehler:disconnected
    isClient		 : BOOL;
    seqNbr       : UINT;
    maxIdleTime_ms  : UDINT;
    lastSendTime_ms : UDINT;

    Com          : DebugIp;
    befiprResp   : msgBefiprRespData;  // the response message from command CMD_BEFIPR

  END_STRUCT;
#pragma pack (pop)

END_TYPE

#define MAX_LOGINS_R             16

VAR_PRIVATE
  rs232Itfs : ARRAY[0..NBR_OF_RS232_ITFS-1] OF RS232_ITF;
  loginArrayR    : ARRAY[0..(MAX_LOGINS_R - 1)] of ^loginContextR;
  loginAnzR      : UDINT;
  comlinkMutexR : MT_SEMAHANDLE;
  comlinkEventR : MT_SEMAHANDLE;
  taskHandleCyclic : UDINT;
  isComlinkRInitialized : BOOL;
  g_lockCnt : UDINT;
  g_inCS : UDINT;
END_VAR

#define LOCK_R()    OS_MT_Wait(comlinkMutexR)
#define UNLOCK_R()  OS_MT_Signal(comlinkMutexR)

FUNCTION ScanL1Block
VAR_INPUT
  pL0Buffer : ^SER_L0_BUF;
  nextOfs : ^UDINT;
  nRead : ^UDINT;
END_VAR
VAR_OUTPUT
  pL1Buffer : ^SER_L1_BUF;
END_VAR;

(*
        SERUSERBAUD_300 (0)
        SERUSERBAUD_600 (1)
        SERUSERBAUD_1200 (2)
        SERUSERBAUD_2400 (3)
        SERUSERBAUD_4800 (4)
        SERUSERBAUD_9600 (5)
        SERUSERBAUD_14400 (6)
        SERUSERBAUD_19200 (7)
        SERUSERBAUD_38400 (8)
        SERUSERBAUD_56000 (9)
        SERUSERBAUD_115200 (10)
*)
FUNCTION GetL0TimeoutValR
VAR_INPUT
  baudrate : UINT;
END_VAR
VAR_OUTPUT
  timeoutVal : UDINT;
END_VAR
VAR
  fact : UDINT;
END_VAR

  CASE baudrate OF
    0:  fact := 384;
    1:  fact := 192;
    2:  fact :=  96;
    3:  fact :=  48;
    4:  fact :=  24;
    5:  fact :=  12;
    6:  fact :=   8;
    7:  fact :=   6;
    8:  fact :=   3;
    9:  fact :=   2;
  ELSE  fact :=   1;
  END_CASE;

  timeoutVal := RS232_L0_TIMEOUT_BAUD115KB * fact + RS232_L0_TIMEOUT_GSMDELAY;

END_FUNCTION

(*
  Errechnet die Byte-Checksumme eines Datenblocks
*)
FUNCTION SerMakeChksum8
VAR_INPUT
  chksumIn : BYTE;
  pData : ^BYTE;
  len : UDINT;
END_VAR
VAR_OUTPUT
  chksumOut : BYTE;
END_VAR
//VAR
//  i : UDINT;
//END_VAR

  chksumOut := chksumIn;
  while(len) do
    chksumOut += pData^;
    pData += 1;
    len -= 1;
  end_while;

//  chksumOut := chksumIn;
//  FOR i := 0 TO len-1 DO
//    chksumOut += pData^;
//    pData += 1;
//  END_FOR;

END_FUNCTION

(*
  Errechnet die Word-Checksumme eines Datenblocks
*)
FUNCTION SerMakeChksum16
VAR_INPUT
  chksumIn : UINT;
  pData : ^BYTE;
  len : UDINT;
END_VAR
VAR_OUTPUT
  chksumOut : UINT;
END_VAR
//VAR
//  i : UDINT;
//END_VAR

  chksumOut := chksumIn;
  while(len) do
    chksumOut += pData^;
    pData += 1;
    len -= 1;
  end_while;

//  chksumOut := chksumIn;
//  FOR i := 0 TO len-1 DO
//    chksumOut += pData^;
//    pData += 1;
//  END_FOR;

END_FUNCTION

(*
  Gibt die Größe eines L0 Pakets in Bytes zurück
*)
FUNCTION GetL0PktLen
VAR_INPUT
  pL0Block : ^SER_L0_BUF;
END_VAR
VAR_OUTPUT
  len : UDINT;
END_VAR

  len := pL0Block^.dataLen + L0_EMPTY_DATALEN;

END_FUNCTION

(*
  Gibt die Größe eines L1 Pakets in Bytes zurück
*)
FUNCTION GetL1PktLen
VAR_INPUT
  pL1Block : ^SER_L1_BUF;
END_VAR
VAR_OUTPUT
  len : UINT;
END_VAR

  len := pL1Block^.dataLen + 5;

END_FUNCTION

(*
  Errechnet die Checksumme eines L0 Blocks
*)
FUNCTION CalcL0DataChksum
VAR_INPUT
  pL0Block : ^SER_L0_BUF;
END_VAR
VAR_OUTPUT
  chksum : UINT;
END_VAR

  chksum := SerMakeChksum16(16#FFFF, #pL0Block^.flagsCmd, GetL0PktLen(pL0Block) - 8);

END_FUNCTION

(*
  Errechnet die Checksumme eines L0 Headers
*)
FUNCTION CalcL0HdrChksum
VAR_INPUT
  pL0Block : ^SER_L0_BUF;
END_VAR
VAR_OUTPUT
  chksum : BYTE;
END_VAR

  chksum := SerMakeChksum8(16#FF, #pL0Block^.dataLen$BYTE, 5);

END_FUNCTION

(*
  Liefert das Cmd-Byte eines L1 Buffers
*)
FUNCTION GetL1CmdR
VAR_INPUT
  pL1Buffer : ^SER_L1_BUF;
END_VAR
VAR_OUTPUT
  cmd : BYTE;
END_VAR

  cmd := pL1Buffer^.flagsCmd AND RS232_L1CMD_MASK;

END_FUNCTION

(*
  Liefert die SeqNbr eines L1 Buffers
*)
FUNCTION GetL1SeqNbrR
VAR_INPUT
  pL1Buffer : ^SER_L1_BUF;
END_VAR
VAR_OUTPUT
  seqNbr : UINT;
END_VAR

  seqNbr := pL1Buffer^.data$UINT;

END_FUNCTION

(*
  Stellt einen L1Block in den L0-Sendebuffer.
  Wenn kein Platz mehr im L0-Sendebuffer ist, dann wird -1 zurückgegeben,
  ansonsten 0.
  Die Checksumme und das ETX Bytes wird hier nicht aktualisiert, das muss am
  Ende gemacht werden, wenn alle L1 Blöcke in den L0 Block gelegt worden sind.
*)
FUNCTION PackL1Block
VAR_INPUT
  pLogin    : ^loginContextR;
  pL1Buffer : ^SER_L1_TXBUF;
END_VAR
VAR_OUTPUT
  retVal : comlinkReason;
END_VAR
VAR
  pL0Buffer : ^SER_L0_BUF;
  l0PktLen : UDINT;
  l1PktLen : UINT;
  pL1BufferTest : ^SER_L1_BUF;
  pReqMsg1 : ^msgUpdCellReqData;
  pReqMsg2 : ^msgUpdCellReqData;
  nextOfs : UDINT;
  nRead : UDINT;
END_VAR

  IF pL1Buffer^.dataValid = 0 THEN
    retVal := COMLINK_ERR_GENERAL;
    RETURN;
  END_IF;

  pL0Buffer := pLogin^.pItf^.pL0SendBufferCollect;

  IF pL1Buffer^.flagsCmd = (CMD_UPDCELL OR RS232_L1FLAGS_IS_REQUEST) THEN
    // Wenn es sich um einen CMD_UPDCELL Request handelt, dann wird der
    // Sendebuffer daraufhin untersucht, ob bereits ein CMD_UPDCELL mit
    // der gleichen LasalID vorhanden ist. Wenn ja, dann werden nur die Daten
    // im Request aktualisiert. Damit wird verhindert, dass der Sendebuffer
    // mit CMD_UPDCELL's von sich rasch ändernden LasalID's überflutet wird.
    nextOfs := SER_L0_BUF.data;
    WHILE nextOfs < (pL0Buffer^.dataLen + 2) DO
      pL1BufferTest := ScanL1Block(pL0Buffer, #nextOfs, #nRead);
      IF pL1BufferTest^.flagsCmd = pL1Buffer^.flagsCmd THEN
        pReqMsg1 := #pL1Buffer^.data[0]$msgUpdCellReqData;
        pReqMsg2 := #pL1BufferTest^.data[0]$msgUpdCellReqData;
        IF (pReqMsg1^.iOff = pReqMsg2^.iOff) & (pReqMsg1^.pCh = pReqMsg2^.pCh) THEN
          // Der Befehl ist gefunden worden -> dData aktualisieren und return
          DEBUGLOG0("%010d-    PackL1Block: data updated in send buffer");
          pReqMsg2^.dData := pReqMsg1^.dData;
          retVal := 0;
          RETURN;
        END_IF;
      END_IF;
    END_WHILE;
  END_IF;

  l0PktLen := GetL0PktLen(pL0Buffer);
  l1PktLen := GetL1PktLen(#pL1Buffer^.srcChIdx$SER_L1_BUF);
  IF (l0PktLen + l1PktLen) > SIZEOF(SER_L0_BUF) THEN
    // kein Platz mehr vorhanden
    DEBUGLOG0("%010d- ***PackL1Block: no more space in send buffer");
    retVal := COMLINK_ERR_GENERAL;
    RETURN;
  END_IF;

  _memcpy(pL0Buffer + l0PktLen - 3, #pL1Buffer^.srcChIdx, l1PktLen);
  pL0Buffer^.dataLen += l1PktLen$UINT;

  // Die Message wurde aus dem Source Buffer in den Transferbuffer kopiert,
  // daher wird dataValid im Source Buffer auf 0 gesetzt.
  pL1Buffer^.dataValid := 0;

  pLogin^.lastSendTime_ms := ops.tAbsolute;

  retVal := 0;

END_FUNCTION

(*
  Errechnet die Checksummen eines L0 Blocks und schreibt die Checksummen
  und das ETX Byte in den L0 Block
*)
FUNCTION FinishL0Block
VAR_INPUT
  pL0Buffer : ^SER_L0_BUF;
END_VAR

  pL0Buffer^.hdrChksum := CalcL0HdrChksum(pL0Buffer);
  (pL0Buffer + GetL0PktLen(pL0Buffer) - 3)$^UINT^ := CalcL0DataChksum(pL0Buffer);
  (pL0Buffer + GetL0PktLen(pL0Buffer) - 1)$^BYTE^ := L0_ETX;

END_FUNCTION

FUNCTION ResetL0
VAR_INPUT
  pItf : ^RS232_ITF;
END_VAR

  _memset(#pItf^.l0SendBufA, 0, SIZEOF(pItf^.l0SendBufA));
  pItf^.l0SendBufA.stx := L0_STX;
  pItf^.l0SendBufA.dataLen := L0_EMPTY_DATALEN;

  _memset(#pItf^.l0SendBufB, 0, SIZEOF(pItf^.l0SendBufB));
  pItf^.l0SendBufB.stx := L0_STX;
  pItf^.l0SendBufB.dataLen := L0_EMPTY_DATALEN;

  pItf^.pL0SendBufferCollect  := #pItf^.l0SendBufA;
  pItf^.pL0SendBufferTransfer := #pItf^.l0SendBufA;
  pItf^.bytesToSend := 0;
  pItf^.bytesSent := 0;
  pItf^.sendInProgress := FALSE;

  pItf^.l0RespPending := FALSE;
  pItf^.l0RespNecessary := FALSE;
  pItf^.l0RespPendingTimeout_ms := pItf^.timeoutVal * 2;
  pItf^.l0RespNecessaryTimeval_ms := RS232_L0_RESP_TIMEVAL;

  pItf^.bytesInRecvBuf := 0;

END_FUNCTION

FUNCTION ResetL1
VAR_INPUT
  pLogin : ^loginContextR;
END_VAR

  pLogin^.isConnected := FALSE;
  pLogin^.hisChIdx := UNKNOWN_CHIDX;
  pLogin^.txL1BufCmd.dataValid := 0;
  pLogin^.txL1BufRefr.dataValid := 0;

END_FUNCTION

//------------------------------------------------------------------------------
// DisconnectAfterErrorR
//  Beendet die Verbindung nachdem ein Fehler festgestellt wurde.
//------------------------------------------------------------------------------
FUNCTION DisconnectAfterErrorR
VAR_INPUT
  pLogin : ^loginContextR;
END_VAR

  DEBUGLOG0("%010d-*** DisconnectAfterErrorR");

  ResetL1(pLogin);

END_FUNCTION

(*
  Beendet alle Verbindungen eines Interfaces
*)
FUNCTION DisconnectAllForItf
VAR_INPUT
  pItf : ^RS232_ITF;
END_VAR
VAR
  i : DINT;
  pLogin : ^loginContextR;
END_VAR

  FOR i := 0 TO (arraysize(loginArrayR) - 1) DO
    pLogin := loginArrayR[i];
    IF pLogin <> NIL & pLogin^.pItf = pItf THEN
      DisconnectAfterErrorR(pLogin);
    END_IF;
  END_FOR;

END_FUNCTION

(*
  Prüft, ob das Senden möglich ist, wenn ja dann wird der L0SendBufferTransfer
  fürs Senden vorbereitet (Flags, Checksumme) und dann wird pItf^.sendInProgress
  auf TRUE gesetzt.

  Es gibt 4 Zustände auf L0 Ebene:
    Resp.Pending  Resp.Necessary  Nächster Send  Kann gesendet werden ?
    ------------  --------------  -------------  ----------------------
    0             0               L0-Request     ja
    1             0               -              nein
    0             1               L0-Response    ja
    1             1               L0-Response    ja
*)
FUNCTION L0CheckSend
VAR_INPUT
  pItf : ^RS232_ITF;
END_VAR

(*
  // Timeouts abfragen und Flags bei abgelaufenen Timeouts berichtigen.
  IF pItf^.l0RespPending & ((ops.tAbsolute - pItf^.l0RespPendingTimeout_ms)$DINT > 0) THEN
    // Es darf nicht ewig auf eine Response gewartet werden.
    DEBUGLOG0("%010d-*** L0CheckSend: timeout for l0RespPending exceeded, resetting connections");
    DisconnectAllForItf(pItf);
    ResetL0(pItf);
    RETURN;
  END_IF;
  *)

  // L0-Sendebuffer ermitteln
  IF pItf^.l0RespPending & !!pItf^.l0RespNecessary THEN
    //DEBUGLOG0("%010d-*** L0CheckSend: send not possible");
    RETURN;
  END_IF;

  IF pItf^.l0RespNecessary THEN
    pItf^.pL0SendBufferTransfer^.flagsCmd  := RS232_L0CMD;
  ELSE
    pItf^.pL0SendBufferTransfer^.flagsCmd  := RS232_L0CMD OR RS232_L0FLAGS_IS_REQUEST;
  END_IF;

  FinishL0Block(pItf^.pL0SendBufferTransfer);

  DEBUGLOG2("%010d-    L0CheckSend: send started, flags: respPending=%d, respNecessary=%d", pItf^.l0RespPending, pItf^.l0RespNecessary);

  pItf^.sendInProgress := TRUE;

END_FUNCTION

(*
  Sendet die Daten im L0SendBufferTransfer.

  Bedingungen:
  Es müssen Daten vorhanden sein und das sendInProgress Flag muss auf TRUE stehen.
*)
FUNCTION L0Send
VAR_INPUT
  pItf : ^RS232_ITF;
END_VAR
VAR
  nWritten : UDINT;
END_VAR

  SERUSER_Send(pItf^.hComm,
               pItf^.pL0SendBufferTransfer + pItf^.bytesSent,
               pItf^.bytesToSend,
               #nWritten);
  pItf^.bytesSent   += nWritten;
  pItf^.bytesToSend -= nWritten;

  DEBUGLOG1("%010d-    L0Send: %d bytes sent", nWritten);

END_FUNCTION

(*
  Liest einen L0-Buffer von der Schnittstelle
*)
FUNCTION L0Recv
VAR_INPUT
  pItf : ^RS232_ITF;
END_VAR
VAR_OUTPUT
  pL0Buffer : ^SER_L0_BUF;
END_VAR
VAR
  bytes2read : UDINT;
  bytesRead : UDINT;
  l0PktLen : UDINT;
  pL0Temp : ^SER_L0_BUF;
  rc : DINT;
END_VAR

  pL0Buffer := NIL;
  pL0Temp := #pItf^.l0RecvBuf$SER_L0_BUF;

  WHILE pItf^.bytesInRecvBuf < SER_L0_BUF.data DO
    bytes2read := (SER_L0_BUF.data)$UDINT - pItf^.bytesInRecvBuf;
    rc := SERUSER_RecvBlock(pItf^.hComm,
                         #pItf^.l0RecvBuf[pItf^.bytesInRecvBuf],
                         bytes2read,
                         #bytesRead);
    IF rc <> 0 THEN
      RETURN;
    END_IF;
    pItf^.bytesInRecvBuf += bytesRead;
    DEBUG_VERBOSE2("%010d-*** L0Recv: %d bytes read, new bytes in recvBuf: %d", bytesRead, pItf^.bytesInRecvBuf);
    IF pItf^.bytesInRecvBuf = SER_L0_BUF.data THEN
      IF (pItf^.l0RecvBuf[0] <> L0_STX) | (CalcL0HdrChksum(pL0Temp) <> pL0Temp^.hdrChksum) THEN
        _memmove(#pItf^.l0RecvBuf[0], #pItf^.l0RecvBuf[1], 6);
        pItf^.bytesInRecvBuf -= bytesRead;
      END_IF;
    END_IF;
  END_WHILE;

  l0PktLen := GetL0PktLen(pL0Temp);
  WHILE pItf^.bytesInRecvBuf < l0PktLen DO
    bytes2read := l0PktLen - pItf^.bytesInRecvBuf;
    rc := SERUSER_RecvBlock(pItf^.hComm,
                            #pItf^.l0RecvBuf[pItf^.bytesInRecvBuf],
                            bytes2read,
                            #bytesRead);
    IF rc <> 0 THEN
      RETURN;
    END_IF;
    pItf^.bytesInRecvBuf += bytesRead;
    DEBUG_VERBOSE2("%010d-*** L0Recv: %d bytes read, new bytes in recvBuf: %d", bytesRead, pItf^.bytesInRecvBuf);
    IF pItf^.bytesInRecvBuf = l0PktLen THEN
      IF (pItf^.l0RecvBuf[l0PktLen-1] = L0_ETX) &
         (CalcL0DataChksum(pL0Temp) = pItf^.l0RecvBuf[l0PktLen-3]$UINT) THEN
        pL0Buffer := pL0Temp;
        IF pL0Temp^.flagsCmd AND RS232_L0FLAGS_IS_REQUEST THEN
          pItf^.l0RespNecessary := TRUE;
        ELSE
          pItf^.l0RespPending := FALSE;
        END_IF;
      END_IF;
      pItf^.bytesInRecvBuf := 0;
      DEBUGLOG2("%010d-    L0Recv: L0 block complete, new flags: respPending=%d, respNecessary=%d", pItf^.l0RespPending, pItf^.l0RespNecessary);
      RETURN;
    END_IF;
  END_WHILE;

END_FUNCTION

(*
  Entnimmt den nächsten L1 Block aus einem L0-Buffer
*)
FUNCTION ScanL1Block
VAR_INPUT
  pL0Buffer : ^SER_L0_BUF;
  nextOfs : ^UDINT;
  nRead : ^UDINT;
END_VAR
VAR_OUTPUT
  pL1Buffer : ^SER_L1_BUF;
END_VAR

  IF nextOfs^ < (pL0Buffer^.dataLen + 3) THEN
    pL1Buffer := pL0Buffer + nextOfs^;
    nRead^ := pL1Buffer^.dataLen + 5;
    nextOfs^ += nRead^;
  ELSE
    nRead^ := 0;
    pL1Buffer := NIL;
  END_IF;

END_FUNCTION

(*
  Liefert einen Zeiger auf den jeweils anderen der beiden Sendebuffer.
*)
FUNCTION SwitchL0Buffer
VAR_INPUT
  pItf : ^RS232_ITF;
  pL0SendBufferIn : ^SER_L0_BUF;
END_VAR
VAR_OUTPUT
  pL0SendBufferOut : ^SER_L0_BUF;
END_VAR

  IF pL0SendBufferIn = #pItf^.l0SendBufA THEN
    pL0SendBufferOut := #pItf^.l0SendBufB;
  ELSE
    pL0SendBufferOut := #pItf^.l0SendBufA;
  END_IF;

END_FUNCTION

//------------------------------------------------------------------------------
// AllocateLoginContextR
//------------------------------------------------------------------------------
FUNCTION AllocateLoginContextR
VAR_INPUT
    interface : UDINT;         // COM Interface number
END_VAR
VAR_OUTPUT
    pLogin       : ^loginContextR;
END_VAR
VAR
    pStatCells  : ^comStCell;
    pDynCells   : ^comStCell;
    mutexName   : ARRAY[0..30] OF CHAR;
END_VAR

  pStatCells := NIL;
  pDynCells  := NIL;

  pLogin := calloc(SIZEOF(loginContextR))$^loginContextR;
  IF pLogin = NIL THEN
    RETURN;
  END_IF;

  // initialize the new connection context
  pStatCells := MemoryUpdateList(#pLogin^.statList, INIT_STATLIST_ENTRIES, 0, 0);
  pDynCells  := MemoryUpdateList(#pLogin^.dynList, INIT_DYNLIST_ENTRIES, 1, 0);
  _strcpy(#mutexName[0], "LOGIN_SEMA_R");
  MakeResourceName(pLogin$UDINT, #mutexName[0]);
  pLogin^.hMutex := OS_MT_CreateSemaphore(MTSEMATYPE_COUNTING,
                                          1,    // initvalue
                                          0,    // flags: 0 means create unconitionally
                                          #mutexName[0]
                                          );
  IF (pStatCells <> NIL) & (pDynCells <> NIL) & (pLogin^.hMutex <> NIL) THEN
    pLogin^.interface  := interface;
    pLogin^.pCallback := g_pCallback;
    pLogin^.hComchMutex := NewComchMutex(pLogin$UDINT, 'r');
    pLogin^.typeOfStruct := STRUCT_TYPE_LOGINCONTEXTR;

    pLogin^.sizeofStatList := MAX_STATLIST_ENTRIES;
    pLogin^.sizeofDynList  := MAX_DYNLIST_ENTRIES;

     // Die Refreshlisten-Größen der Remote Station werden vorerst mit der Größe der eigenen
     // initialisiert. Wenn beim Login ein anderer Wert gemeldet wird, dann wird diese
     // Variable noch einmal überschrieben
    pLogin^.sizeofRemoteDynList  := pLogin^.sizeofDynList;
    pLogin^.sizeofRemoteStatList := pLogin^.sizeofStatList;

    pLogin^.hisChIdx := INVALID_CHIDX;

    DEBUGLOG0("%010d-  =====  Login context allocated  =====");
  ELSE
    // cleanup
    IF pLogin^.hMutex <> NIL THEN
      OS_MT_DeleteSemaphore(pLogin^.hMutex);
    END_IF;
    IF pStatCells <> NIL THEN
      _free(pStatCells);
      pStatCells := NIL;
      g_nbrStatList -= 1;
    END_IF;
    IF pDynCells <> NIL THEN
      _free(pDynCells);
      pDynCells := NIL;
      g_nbrDynList -= 1;
    END_IF;
    _free(pLogin);
    pLogin := NIL;
  END_IF;

END_FUNCTION

//------------------------------------------------------------------------------
// ReleaseLoginContextR
//
//  Release all resources of a used login context.
//------------------------------------------------------------------------------
FUNCTION ReleaseLoginContextR
VAR_INPUT
    pLogin       : ^loginContextR;
END_VAR

  IF pLogin = NIL THEN
    RETURN;
  END_IF;

  IF pLogin^.hMutex <> NIL THEN
    OS_MT_DeleteSemaphore(pLogin^.hMutex);
  END_IF;
  DeleteComchMutex(#pLogin^.hComchMutex);

  IF pLogin^.pNode <> NIL THEN
    RemoveMonitorNode(pLogin^.pNode);
  END_IF;

  IF pLogin^.pComdefT THEN
    pLogin^.pComdefT^.pLogin := NIL;
  END_IF;

  // free allocated memory
  _free(pLogin^.statList.pFirstCell);
  g_nbrStatList -= 1;
  _free(pLogin^.dynList.pFirstCell);
  g_nbrDynList -= 1;
  pLogin^.statList.pFirstCell := NIL;
  pLogin^.dynList.pFirstCell := NIL;

  _free(pLogin);
  pLogin := NIL;

  DEBUGLOG0("%010d-  =====  Login context released  =====");

END_FUNCTION

(*
  Wandelt eine Interface Nummer (in ComTypes.h definiert, z.B.COMLINK_IFNUM_COM1)
  in einen Interface Index um. Dieser Index kann für das Array rs232Itfs verwendet
  werden.
  Bei einem Fehler wird -1 zurückgegeben.
*)
FUNCTION ComlinkR_Itfnbr2Idx
VAR_INPUT
  interface : UDINT;
END_VAR
VAR_OUTPUT
  idx : DINT;
END_VAR

  CASE interface OF
    COMLINK_IFNUM_COM1,
    COMLINK_IFNUM_COM2,
    COMLINK_IFNUM_COM3,
    COMLINK_IFNUM_COM4:
      idx$UDINT := interface - COMLINK_IFNUM_COM1;
    COMLINK_IFNUM_COM5,
    COMLINK_IFNUM_COM6,
    COMLINK_IFNUM_COM7,
    COMLINK_IFNUM_COM8,
    COMLINK_IFNUM_COM9,
    COMLINK_IFNUM_COM10:
      idx$UDINT := interface - COMLINK_IFNUM_COM5 + 4;
    ELSE
      idx := -1;
  END_CASE;

  IF idx >= arraysize(rs232Itfs) THEN
    idx := -1;
  END_IF;

END_FUNCTION

(*
  Wandelt einen Interface Index in eine Interface Nummer (in ComTypes.h definiert,
  z.B.COMLINK_IFNUM_COM1) um.
*)
FUNCTION ComlinkR_Idx2Itfnbr
VAR_INPUT
  idx : DINT;
END_VAR
VAR_OUTPUT
  interface : UDINT;
END_VAR

  IF idx < 4 THEN
    interface := idx$UDINT + COMLINK_IFNUM_COM1;
  ELSE
    interface := idx$UDINT + COMLINK_IFNUM_COM5;
  END_IF;

END_FUNCTION

//------------------------------------------------------------------------------
// ComlinkR_GetHandle
//  Gibt das zu einer Interface Nummmer gehörende Handle zurück.
//  Wenn es nocht nicht initialisiert worden ist, dann wird das hier gemacht.
//------------------------------------------------------------------------------
FUNCTION ComlinkR_GetHandle
VAR_INPUT
  interface : UDINT;
END_VAR
VAR_OUTPUT
  hComm : pVoid;
END_VAR
VAR
  idx : DINT;
  pItf : ^RS232_ITF;
  initStatus : DINT;
END_VAR

  idx := ComlinkR_Itfnbr2Idx(interface);

  IF idx >= 0 THEN
    pItf := #rs232Itfs[idx];
    hComm := pItf^.hComm;
    IF hComm = NIL THEN
      IF pItf^.hCommAppl = NIL THEN
        pItf^.hCommAppl := SERUSER_Init(idx$UINT + 1, pItf^.baudrate, DFLT_PARITY, DFLT_STOP, DFLT_WORDL);
      END_IF;
      IF pItf^.hCommAppl <> NIL THEN
        g_RS232activity := TRUE;

        IF pItf^.fnInitInterface <> NIL THEN
          initStatus := pItf^.fnInitInterface$LDR_InitRs232Interface(pItf^.pThis, interface, pItf^.hCommAppl);
        ELSE
          initStatus := 1;
        END_IF;
        IF initStatus > 0 THEN
          hComm := pItf^.hCommAppl;
          pItf^.hComm := hComm;
        END_IF;
      END_IF;
    END_IF;
  ELSE
    hComm := NIL;
  END_IF;

END_FUNCTION

//------------------------------------------------------------------------------
// ComlinkR_Init
//------------------------------------------------------------------------------
FUNCTION ComlinkR_Init
VAR
  i : DINT;
END_VAR

  IF mt_api = NIL | _LSL_POS^.piSSR^.SSR_CurrentTaskHandle = NIL THEN
    isComlinkRInitialized := FALSE;
    RETURN;
  END_IF;

  _memset(#rs232Itfs[0], 0, SIZEOF(rs232Itfs));
  FOR i := 0 TO arraysize(rs232Itfs)-1 DO
    rs232Itfs[i].itfIdx := i;
    rs232Itfs[i].baudrate := DFLT_BAUD;
    rs232Itfs[i].timeoutVal := GetL0TimeoutValR(rs232Itfs[i].baudrate);
    ResetL0(#rs232Itfs[i]);
    DEBUGLOG2("%010d-    ComlinkR_Init: itf %d - timeoutVal=%d", i$UDINT, rs232Itfs[i].timeoutVal);
  END_FOR;

  _memset(#loginArrayR[0], 0, SIZEOF(loginArrayR));
  loginAnzR         := 0;

  comlinkMutexR := OS_MT_CreateSemaphore(MTSEMATYPE_MUTEX,
                                         1,    // initvalue
                                         0,    // flags: 0 means create unconitionally
                                         "COMLINKR_MUTEX0"
                                         );
  comlinkEventR := OS_MT_CreateSemaphore(MTSEMATYPE_EVENT,
                                         0,    // initvalue
                                         0,    // flags: 0 means create unconitionally
                                         "COMLINKR_EVENT0"
                                         );

  taskHandleCyclic := OS_SSR_CurrentTaskHandle();

  isComlinkRInitialized := TRUE;

END_FUNCTION

(*
  Blockiert so lange, bis eine RS232 Übertragung stattgefunden hat.

  Wenn der Aufruf ausserhalb des Cyclic erfolgt, dann blockiert diese Funktion
  auf einem Event Semaphore, das vom Cyclic in der ComlinkR_SerTransfer Funktion
  gepulst wird.

  Wenn der Aufruf im Context des Cyclic Tasks erfolgt, dann muss die ComlinkR_SerTransfer
  Funktion selbst aufgerufen werden, weil ja der Loader-Cyclic nicht aufgerufen
  wird, solange man sich in der RS232WaitForTransfer Funktion befindet.
*)
FUNCTION RS232WaitForTransfer
VAR_INPUT
  pItf : ^RS232_ITF;
END_VAR
VAR
  startTime : UDINT;
END_VAR

  IF OS_SSR_CurrentTaskHandle() = taskHandleCyclic THEN
    startTime := ops.tAbsolute;
    WHILE (ops.tAbsolute - startTime) < 20 DO
      IF ComlinkR_SerTransfer(pItf) THEN
        RETURN;
      END_IF;
      OS_MT_Delay(1);
    END_WHILE;
  ELSE
    OS_MT_WaitTimed(comlinkEventR, 20);
  END_IF;

END_FUNCTION

//------------------------------------------------------------------------------
// SendRequestR
//  Sendet einen Request
//------------------------------------------------------------------------------
FUNCTION SendRequestR
VAR_INPUT
  pLogin : ^loginContextR;
  cmd : BYTE;
  respRequired : BOOL;
  pData : pVoid;
  dataLen : UDINT;
  blockingMode : BOOL;
END_VAR
VAR_OUTPUT
  retval        : comlinkReason;
END_VAR
VAR
  startTime : UDINT;
  pTxL1Buf : ^SER_L1_TXBUF;
  seqNbrSize : UINT;
END_VAR

  retval := 0;

  IF pLogin^.isConnected = FALSE & pLogin^.hisChIdx <> UNKNOWN_CHIDX THEN
    DEBUGLOG0("%010d-*** SendRequestR: COMLINK_ERR_NOCONNECTION");
    retval := COMLINK_ERR_NOCONNECTION;
    RETURN;
  END_IF;

  IF respRequired THEN
    seqNbrSize := SIZEOF(UINT);
  ELSE
    seqNbrSize := 0;
  END_IF;
  IF dataLen > SIZEOF(pTxL1Buf^.data) - seqNbrSize THEN
    DEBUGLOG0("%010d-*** SendRequestR: COMLINK_ERR_BUF_TOO_SMALL");
    retval := COMLINK_ERR_BUF_TOO_SMALL;
    RETURN;
  END_IF;

  IF respRequired THEN
    pTxL1Buf := #pLogin^.txL1BufCmd;
  ELSE
    pTxL1Buf := #pLogin^.txL1BufRefr;
  END_IF;

  pTxL1Buf^.srcChIdx := pLogin^.myChIdx;
  pTxL1Buf^.dstChIdx := pLogin^.hisChIdx;
  pTxL1Buf^.flagsCmd := cmd OR RS232_L1FLAGS_IS_REQUEST;

  IF respRequired THEN
    pLogin^.seqNbr += 1;
    pTxL1Buf^.flagsCmd := pTxL1Buf^.flagsCmd OR RS232_L1FLAGS_RESPONSE_REQUIRED;
    pTxL1Buf^.dataLen  := SIZEOF(UINT);
    pTxL1Buf^.data$UINT := pLogin^.seqNbr;
    // Wenn srcChIdx im L1 RxBuffer auf INVALID_CHIDX gesetzt wird, dann heisst das,
    // dass der Buffer leer ist und vom Übertragungsteil beschrieben werden darf.
    pLogin^.rxL1BufResp.srcChIdx := INVALID_CHIDX;
  ELSE
    pTxL1Buf^.dataLen := 0;
  END_IF;

  _memcpy(#pTxL1Buf^.data[0] + pTxL1Buf^.dataLen, pData, dataLen);
  pTxL1Buf^.dataLen += dataLen$UINT;

  pTxL1Buf^.dataValid := 1;

  startTime := OPS.tAbsolute;
  WHILE 1 DO
    LOCK_R();
    retval := PackL1Block(pLogin, pTxL1Buf);
    UNLOCK_R();
    IF retval = 0 THEN
      IF respRequired THEN
        DEBUGLOG3("%010d- 1> ch%d SendRequestR: put L1 message into collect buffer: dataLen(incl.seqNbr)=%d, seqNbr=%d", pLogin^.myChIdx, pTxL1Buf^.dataLen, TO_UDINT(pTxL1Buf^.data$UINT));
      ELSE
        DEBUGLOG2("%010d- 1> ch%d SendRequestR: put L1 message into collect buffer: dataLen=%d", pLogin^.myChIdx, pTxL1Buf^.dataLen);
      END_IF;
      EXIT;
    END_IF;

    IF !!blockingMode THEN
      EXIT;
    END_IF;

    IF (OPS.tAbsolute - startTime) > pLogin^.pItf^.timeoutVal THEN
      DEBUGLOG0("%010d-*** SendRequestR: COMLINK_ERR_TIMEOUT");
      retval := COMLINK_ERR_TIMEOUT;
      EXIT;
    END_IF;

    RS232WaitForTransfer(pLogin^.pItf);

  END_WHILE;

  pTxL1Buf^.dataValid := 0;

END_FUNCTION

//------------------------------------------------------------------------------
// WaitForResponseR
//  Wartet auf die Response
//------------------------------------------------------------------------------
FUNCTION WaitForResponseR
VAR_INPUT
  pLogin : ^loginContextR;
  pRespData : pVoid;
  respDataLen : UINT;
END_VAR
VAR_OUTPUT
  retval        : INT;
END_VAR
VAR
  startTime : UDINT;
END_VAR

  IF pLogin^.isConnected = FALSE & pLogin^.hisChIdx <> UNKNOWN_CHIDX THEN
    DEBUGLOG0("%010d-*** WaitForResponseR: COMLINK_ERR_NOCONNECTION");
    retval := COMLINK_ERR_NOCONNECTION$INT;
    RETURN;
  END_IF;

  startTime := OPS.tAbsolute;
  WHILE 1 DO
    IF (pLogin^.rxL1BufResp.srcChIdx <> INVALID_CHIDX) THEN
      IF ((pLogin^.rxL1BufResp.flagsCmd$USINT AND RS232_L1CMD_MASK) = (pLogin^.txL1BufCmd.flagsCmd$USINT AND RS232_L1CMD_MASK)) THEN
        IF (pLogin^.rxL1BufResp.dataLen >= SIZEOF(UINT)) THEN
          IF (pLogin^.rxL1BufResp.data$UINT = pLogin^.seqNbr) THEN

            DEBUGLOG3("%010d-<1  ch%d WaitForResponseR: received expected L1 message: dataLen(incl.seqNbr)=%d, seqNbr=%d", pLogin^.myChIdx, pLogin^.rxL1BufResp.dataLen, TO_UDINT(pLogin^.seqNbr));
            IF pLogin^.rxL1BufResp.flagsCmd AND RS232_L1FLAGS_ACK THEN
              retval := 0;
              IF respDataLen > pLogin^.rxL1BufResp.dataLen - SIZEOF(UINT) THEN
                respDataLen := pLogin^.rxL1BufResp.dataLen - SIZEOF(UINT);
              END_IF;
              IF pRespData <> NIL THEN
                _memcpy(pRespData, #pLogin^.rxL1BufResp.data[2], respDataLen);
              END_IF;
              retval := respDataLen$INT;
            ELSE
              DEBUGLOG0("%010d-*** WaitForResponseR: COMLINK_ERR_INVALID_RESPONSE");
              retval := COMLINK_ERR_INVALID_RESPONSE$INT;
            END_IF;
            EXIT;

          ELSE
            DEBUGLOG2("%010d-*** WaitForResponseR: received unexpected L1 message, rcvdSeqNbr=%d, expctdSeqNbr=%d", TO_UDINT(pLogin^.rxL1BufResp.data$UINT), TO_UDINT(pLogin^.seqNbr));
          END_IF;
        ELSE
          DEBUGLOG1("%010d-*** WaitForResponseR: received unexpected L1 message, invalid dataLen=%d", TO_UDINT(pLogin^.rxL1BufResp.dataLen));
        END_IF;
      ELSE
        DEBUGLOG2("%010d-*** WaitForResponseR: received unexpected L1 message, rcvdCmd=%d, expctdCmd=%d", TO_UDINT(pLogin^.rxL1BufResp.flagsCmd$USINT AND RS232_L1CMD_MASK), TO_UDINT(pLogin^.txL1BufCmd.flagsCmd$USINT AND RS232_L1CMD_MASK));
      END_IF;
    END_IF;

    IF (OPS.tAbsolute - startTime) > pLogin^.pItf^.timeoutVal THEN
      DEBUGLOG1("%010d-*** ch%d WaitForResponseR: COMLINK_ERR_TIMEOUT", pLogin^.myChIdx);
      retval := COMLINK_ERR_TIMEOUT$INT;
      EXIT;
    END_IF;

    RS232WaitForTransfer(pLogin^.pItf);

  END_WHILE;

END_FUNCTION

//------------------------------------------------------------------------------
// SendResponseR
//  Sendet eine Response
//------------------------------------------------------------------------------
FUNCTION SendResponseR
VAR_INPUT
  pLogin : ^loginContextR;
  seqNbr : UINT;
  ack : BOOL;
  cmd : BYTE;
  pData : pVoid;
  dataLen : UDINT;
END_VAR
VAR_OUTPUT
  retval        : comlinkReason;
END_VAR
VAR
  pTxL1Buf : ^SER_L1_TXBUF;
END_VAR

  retval := 0;

  IF sizeof(UINT) + dataLen > SIZEOF(pTxL1Buf^.data) THEN
    DEBUGLOG0("%010d-*** SendResponseR: COMLINK_ERR_BUF_TOO_SMALL");
    retval := COMLINK_ERR_BUF_TOO_SMALL;
    RETURN;
  END_IF;

  pTxL1Buf := #pLogin^.txL1BufCmd;

  IF pTxL1Buf^.dataValid THEN
    DEBUGLOG0("%010d-*** SendResponseR: txBuf is not free");
    retval := COMLINK_ERR_BUF_TOO_SMALL;
    RETURN;
  END_IF;

  pTxL1Buf^.srcChIdx := pLogin^.myChIdx;
  pTxL1Buf^.dstChIdx := pLogin^.hisChIdx;
  pTxL1Buf^.flagsCmd := cmd AND RS232_L1CMD_MASK;
  IF ack THEN
    pTxL1Buf^.flagsCmd := pTxL1Buf^.flagsCmd OR RS232_L1FLAGS_ACK;
  END_IF;

  pTxL1Buf^.dataLen  := sizeof(UINT) + dataLen$UINT;
  pTxL1Buf^.data$UINT := seqNbr;
  _memcpy(#pTxL1Buf^.data[2], pData, dataLen);

  pTxL1Buf^.dataValid := 1;

  LOCK_R();
  retval := PackL1Block(pLogin, #pTxL1Buf^);
  UNLOCK_R();

  IF retval = 0 THEN
    DEBUGLOG2("%010d- 1> SendResponseR: put L1 message into collect buffer: dataLen(incl.seqNbr)=%d, seqNbr=%d", pTxL1Buf^.dataLen, TO_UDINT(pTxL1Buf^.data$UINT));
  ELSE
    DEBUGLOG2("%010d- 1> *** SendResponseR: PackL1Block failed: dataLen(incl.seqNbr)=%d, seqNbr=%d", pTxL1Buf^.dataLen, TO_UDINT(pTxL1Buf^.data$UINT));
  END_IF;

END_FUNCTION

//------------------------------------------------------------------------------
// ConnectR
//  Schickt den Login Befehl
//------------------------------------------------------------------------------
FUNCTION ConnectR
VAR_INPUT
  pLogin : ^loginContextR;
END_VAR
VAR_OUTPUT
  retval        : DINT;
END_VAR

  ResetL1(pLogin);

  // Request senden
  retval := SendRequestR(pLogin, CMD_CONNECT, respRequired:=TRUE, pData:=NIL, dataLen:=0, blockingMode:=TRUE);
  IF retval <> 0 THEN
    RETURN;
  END_IF;

  // warten auf die Antwort
  retval := WaitForResponseR(pLogin, NIL, 0);
  IF retval >= 0 THEN
    pLogin^.hisChIdx := pLogin^.rxL1BufResp.srcChIdx;
    pLogin^.isConnected := TRUE;
  END_IF;

END_FUNCTION

//------------------------------------------------------------------------------
// ExchgSessionInfoR
//  Exchange session info with the server
//------------------------------------------------------------------------------
FUNCTION ExchgSessionInfoR
VAR_INPUT
  pLogin : ^loginContextR;
  mySessId      : UDINT;
  versionOfPeer : ^UDINT;
  instIdOfPeer  : ^UDINT;
  sizeofRemoteDynList  : ^UINT;
  sizeofRemoteStatList : ^UINT;
END_VAR
VAR_OUTPUT
  retval        : DINT;
END_VAR
VAR
  msgData          : msgSessInfoData;
END_VAR

  msgData.version := COMLINKR_VERSION;
  msgData.instId  := myInstanceId;
  msgData.sessId  := mySessId;
  msgData.sizeofDynList  := MAX_DYNLIST_ENTRIES;
  msgData.sizeofStatList := MAX_STATLIST_ENTRIES;

  // Request senden
  retval := SendRequestR(pLogin,
                         CMD_SESSINFO,
                         respRequired:=TRUE,
                         #msgData,
                         SIZEOF(msgData),
                         blockingMode:=TRUE);
  IF retval <> 0 THEN
    RETURN;
  END_IF;

  // warten auf die Antwort
  retval := WaitForResponseR(pLogin, #msgData, SIZEOF(msgData));
  IF retval >= 0 THEN
    versionOfPeer^:= msgData.version;
    instIdOfPeer^ := msgData.instId;
    sizeofRemoteDynList^  := msgData.sizeofDynList;
    sizeofRemoteStatList^ := msgData.sizeofStatList;
  END_IF;

END_FUNCTION

//------------------------------------------------------------------------------
// IsConnectedR
//  Prüft, ob eine Verbindung besteht. Eine Verbindung ist aufrecht vom Login
//  bis zu einem Fehler. Nach einem Fehler muss wieder ein Login gemacht werden.
//  Beim Login wird der Verbindungsstatus resettiert (z.B. alle Zellen in der
//  Refreshliste auf 0 gesetzt)
//------------------------------------------------------------------------------
FUNCTION IsConnectedR
VAR_INPUT
  pLogin : ^loginContextR;
END_VAR
VAR_OUTPUT
  retval : BOOL;
END_VAR

  retval := pLogin^.isConnected;

END_FUNCTION

//------------------------------------------------------------------------------
// SearchUsedConnBlockCltR
//  Sucht einen vom Client bereits benutzten Connection Block
//------------------------------------------------------------------------------
FUNCTION SearchUsedConnBlockCltR
VAR_INPUT
  pComdef : ^comdef;
END_VAR
VAR_OUTPUT
  pLogin : ^loginContextR; // connection context
END_VAR
VAR
  i : UDINT;
END_VAR

  pLogin := NIL;
  FOR i := 0 TO (arraysize(loginArrayR) - 1) DO
    IF (loginArrayR[i] <> NIL) &
       (loginArrayR[i]^.interface = pComdef^.interface) &
       (loginArrayR[i]^.pComdefT = pComdef$^comdefT) THEN
      pLogin := loginArrayR[i];
      IF pLogin^.pItf^.hComm = 0 THEN
        // ComlinkR_GetHandle erneut aufrufen, damit die Callbackfunktion aufgerufen
        // werden kann.
        pLogin^.pItf^.hComm := ComlinkR_GetHandle(ComlinkR_Idx2Itfnbr(pLogin^.pItf^.itfIdx));
      END_IF;
      IF pLogin^.pItf^.hComm = 0 THEN
        pLogin := NIL;
      END_IF;
      EXIT;
    END_IF;
  END_FOR;

END_FUNCTION

//------------------------------------------------------------------------------
// SearchUsedConnBlockSvrR
//  Sucht einen vom Server bereits benutzten Connection Block
//------------------------------------------------------------------------------
FUNCTION SearchUsedConnBlockSvrR
VAR_INPUT
  itfIdx : DINT;
  remoteChIdx : BYTE;
END_VAR
VAR_OUTPUT
  pLogin : ^loginContextR; // connection context
END_VAR
VAR
  i : UDINT;
END_VAR

  pLogin := NIL;
  FOR i := 0 TO (arraysize(loginArrayR) - 1) DO
    IF (loginArrayR[i] <> NIL) &
       (ComlinkR_Itfnbr2Idx(loginArrayR[i]^.interface) = itfIdx) &
       (loginArrayR[i]^.hisChIdx = remoteChIdx) THEN
      pLogin := loginArrayR[i];
      EXIT;
    END_IF;
  END_FOR;

END_FUNCTION

//------------------------------------------------------------------------------
// AllocNewConnBlockCltR
//  Alloziert für den Client einen neuen Connection Block
//------------------------------------------------------------------------------
FUNCTION AllocNewConnBlockCltR
VAR_INPUT
  pComdefT : ^comdefT;
  pRetval : ^UINT;
END_VAR
VAR_OUTPUT
  pLogin : ^loginContextR; // connection context
END_VAR
VAR
  i : UDINT;
  hComm : pVoid;
END_VAR

  pLogin := NIL;
  IF loginAnzR = arraysize(loginArrayR) THEN
    DEBUGLOG0("%010d-*** AllocNewConnBlockCltR: COMLINK_ERR_MAXCONN");
    pRetval^ := COMLINK_ERR_MAXCONN;
    RETURN;
  END_IF;

  hComm := ComlinkR_GetHandle(pComdefT^.interface);
  IF hComm = 0 THEN
    DEBUGLOG0("%010d-*** AllocNewConnBlockCltR: ComlinkR_GetHandle failed");
    RETURN;
  END_IF;

  // try to get a connection context
  pLogin := AllocateLoginContextR(pComdefT^.interface);
  IF pLogin = NIL THEN
    DEBUGLOG0("%010d-*** AllocNewConnBlockCltR: AllocateLoginContextR failed");
    RETURN;
  END_IF;

  pLogin^.pItf := #rs232Itfs[ComlinkR_Itfnbr2Idx(pComdefT^.interface)];
  pLogin^.pItf^.hComm := hComm;

  // success: try to put pLogin into loginArrayR
  LOCK_R();

  // search a free entry in loginArrayR
  FOR i := 0 TO (arraysize(loginArrayR) - 1) DO
    IF loginArrayR[i] = NIL THEN
      EXIT;
    END_IF;
  END_FOR;
  IF i = arraysize(loginArrayR) THEN
    pRetval^ := COMLINK_ERR_MAXCONN;
    UNLOCK_R();
    ReleaseLoginContextR(pLogin);
    RETURN;
  END_IF;

  pComdefT^.pLogin := pLogin$^loginContext;
  // make an entry in the loginArrayR
  loginArrayR[i] := pLogin;
  pLogin^.myChIdx := i;
  loginAnzR += 1;

  UNLOCK_R();

END_FUNCTION

//------------------------------------------------------------------------------
// AllocNewConnBlockSvrR
//  Alloziert für den Server einen neuen Connection Block
//------------------------------------------------------------------------------
FUNCTION AllocNewConnBlockSvrR
VAR_INPUT
  itfIdx : DINT;
  remoteChIdx : BYTE;
END_VAR
VAR_OUTPUT
  pLogin : ^loginContextR; // connection context
END_VAR
VAR
  i : UDINT;
  interface : UDINT;
END_VAR

  interface := ComlinkR_Idx2Itfnbr(itfIdx);

  pLogin := NIL;
  IF loginAnzR = arraysize(loginArrayR) THEN
    DEBUGLOG0("%010d-*** AllocNewConnBlockSvrR: COMLINK_ERR_MAXCONN");
    RETURN;
  END_IF;

  // try to get a connection context
  pLogin := AllocateLoginContextR(interface);
  IF pLogin = NIL THEN
    DEBUGLOG0("%010d-*** AllocNewConnBlockSvrR: AllocateLoginContextR failed");
    RETURN;
  END_IF;
  pLogin^.pItf := #rs232Itfs[itfIdx];

  pLogin^.pItf^.hComm := ComlinkR_GetHandle(interface);
  IF pLogin^.pItf^.hComm = 0 THEN
    DEBUGLOG0("%010d-*** AllocNewConnBlockSvrR: ComlinkR_GetHandle failed");
    ReleaseLoginContextR(pLogin);
    RETURN;
  END_IF;

  // success: try to put pLogin into loginArrayR
  LOCK_R();

  // search a free entry in loginArrayR
  FOR i := 0 TO (arraysize(loginArrayR) - 1) DO
    IF loginArrayR[i] = NIL THEN
      EXIT;
    END_IF;
  END_FOR;
  IF i = arraysize(loginArrayR) THEN
    UNLOCK_R();
    ReleaseLoginContextR(pLogin);
    RETURN;
  END_IF;

  // make an entry in the loginArrayR
  loginArrayR[i] := pLogin;
  pLogin^.myChIdx := i;
  loginAnzR += 1;

  UNLOCK_R();

END_FUNCTION

FUNCTION ComlinkR_Logout
VAR_INPUT
  pComdef : ^comdef;
END_VAR
VAR_OUTPUT
  retval : UINT;
END_VAR
VAR
  pComDefT : ^comdefT;
END_VAR

  pComDefT := pComdef$^comdefT;
  ReleaseLoginContextR( pComDefT^.pLogin$^loginContextR );
  Seruser_Close( ComlinkR_GetHandle( pComDefT^.Interface ) );
  retval := 0;

END_FUNCTION

//------------------------------------------------------------------------------
// ComlinkR_Login
//  Login über RS232
//------------------------------------------------------------------------------
FUNCTION ComlinkR_Login
VAR_INPUT
    pComdef       : ^comdef;
END_VAR
VAR_OUTPUT
    retval        : UINT;
END_VAR
VAR
    pComdefT      : ^comdefT;
    pLogin        : ^loginContextR; // connection context
    versionOfPeer : UDINT;
    instIdOfPeer  : UDINT;
    rc            : DINT;
    sizeofRemoteDynList  : UINT;
    sizeofRemoteStatList : UINT;
END_VAR

  DEBUGLOG0("%010d-ComlinkR_Login");

  retval   := COMLINK_ERR_GENERAL;

  IF !!isComlinkRInitialized THEN
    RETURN;
  END_IF;

  pComdefT := pComdef$^comdefT;

  pLogin := SearchUsedConnBlockCltR(pComdef);
  IF pLogin = NIL THEN
    pLogin := AllocNewConnBlockCltR(pComdefT, #retval);
  END_IF;

  IF pLogin = NIL THEN
    RETURN;
  END_IF;

  pLogin^.isClient := TRUE;

  //ResetL0(pLogin^.pItf);

  rc := ConnectR(pLogin);
  IF rc <> 0 THEN
    DEBUGLOG1("%010d-*** ComlinkR_Login: ConnectR failed, rc=%d", TO_UDINT(rc));
    retval := rc$UINT;
    RETURN;
  END_IF;

  // exchange session info with the server
  sizeofRemoteDynList  := pLogin^.sizeofRemoteDynList;
  sizeofRemoteStatList := pLogin^.sizeofRemoteStatList;
  rc := ExchgSessionInfoR(pLogin,
                          pComdef$UDINT,
                          #versionOfPeer,
                          #instIdOfPeer,
                          #sizeofRemoteDynList,
                          #sizeofRemoteStatList);
  IF rc < 0 THEN
    DEBUGLOG1("%010d-*** ComlinkR_Login: ExchgSessionInfo failed, rc=%d", TO_UDINT(rc));
    retval := COMLINK_ERR_NOCONNECTION;
    RETURN;
  END_IF;

  retval := 0;
  pLogin^.versionOfPeer := versionOfPeer;
  pLogin^.instIdOfPeer  := instIdOfPeer;
  pLogin^.sizeofRemoteDynList  := sizeofRemoteDynList;
  pLogin^.sizeofRemoteStatList := sizeofRemoteStatList;
  pLogin^.pComdefT      := pComdefT; // this pointer is needed when the callback function is called

END_FUNCTION

//------------------------------------------------------------------------------
// ComlinkR_TxCommandEx
//
//  This function send interpreter code to the comlink server. The server
//  executes the code and responds with the the result and the workstate.
//------------------------------------------------------------------------------
FUNCTION ComlinkR_TxCommandEx
VAR_INPUT
    opCode    : UDINT;
    length    : UDINT;
    aPara     : ^USINT;
    pComdef   : ^comdef;
    pResu     : ^UDINT;
    pStatus   : ^IPRSTATES;
    res       : UDINT;
END_VAR
VAR_OUTPUT
    retval    : comlinkReason;
END_VAR
VAR
    pComdefT  : ^comdefT;
    pLogin    : ^loginContextR; // connection context
    reqMsg    : msgBefiprReqData; // request structure for command CMD_BEFIPR
    reqMsgLen : UDINT;
    fOk       : UDINT;
    rc        : DINT;
END_VAR

  pComdefT := pComdef$^comdefT;
  pStatus^ := ERROR;
  retval   := COMLINK_ERR_GENERAL;
  fOk   := 0;

  IF !!isComlinkRInitialized THEN
    DEBUGLOG0("%010d-*** ComlinkT_TxCommandEx: !!isComlinkRInitialized");
    RETURN;
  END_IF;

  pLogin := pComdefT^.pLogin$^loginContextR;
  IF pLogin = NIL THEN
    DEBUGLOG0("%010d-*** ComlinkT_TxCommandEx: COMLINK_ERR_LOGIN_REQUIRED");
    retval := COMLINK_ERR_LOGIN_REQUIRED;
    RETURN;
  END_IF;

  pResu^ := (#pLogin^.befiprResp.resu)$UDINT;

  IF length > SIZEOF(reqMsg.instr.aPara) THEN
    // parameter length is too big
    DEBUGLOG0("%010d-*** ComlinkT_TxCommandEx: parameter length is too big");
    retval := COMLINK_ERR_INVALID_PARAM;
    RETURN;
  END_IF;

  // prepare the request message structure
  reqMsg.workState    := BUSY;
  reqMsg.instr.opCode := opCode$INSTRSET;
  reqMsg.instr.uiLng  := (length + SIZEOF(instruct.uiLng))$UINT;
  _memcpy(#reqMsg.instr.aPara, aPara, length);

  reqMsgLen := SIZEOF(reqMsg.workState)    +
               SIZEOF(reqMsg.instr.opCode) +
               SIZEOF(reqMsg.instr.uiLng)  +
               length;

  // Send the request
  rc := SendRequestR(pLogin,
                     CMD_BEFIPR,
                     respRequired:=TRUE,
                     #reqMsg,
                     reqMsgLen,
                     blockingMode:=TRUE);
  IF rc <> 0 THEN
    DEBUGLOG1("%010d-*** ComlinkR_TxCommandEx: SendRequestR failed, rc=%d", TO_UDINT(rc));
    retval := COMLINK_ERR_NOCONNECTION;
    GOTO EndLabel;
  END_IF;
  DEBUGLOG2("%010d-ComlinkR_TxCommandEx: BEFIPR request sent, opCode=%d, msgLen=%d", opCode, TO_UDINT(rc));

  // Read the response
  rc := WaitForResponseR(pLogin, #pLogin^.befiprResp, SIZEOF(pLogin^.befiprResp));
  IF rc < 0 THEN
    DEBUGLOG1("%010d-*** ComlinkR_TxCommandEx: ReadCmdMsg failed, rc=%d", TO_UDINT(rc));
    retval := COMLINK_ERR_NOCONNECTION;
    GOTO EndLabel;
  END_IF;
  AliveCheckMsgRcvd(pLogin$^loginContext);

  IF rc < SIZEOF(pLogin^.befiprResp.workstate) THEN
    // not enough data received !
    DEBUGLOG0("%010d-*** ComlinkR_TxCommandEx: not enough data received");
    retval := COMLINK_ERR_INVALID_RESPONSE;
    GOTO EndLabel;
  END_IF;

  fOk := 1;

EndLabel:
  IF fOk = 0 THEN
    // The connection has to be closed because it's possible that partial data
    // is transferred.
    DEBUGLOG0("%010d-ComlinkR_TxCommandEx: closing connection");
    DisconnectAfterErrorR(pLogin);
    pStatus^ := ERROR;
  ELSE
    pStatus^ := pLogin^.befiprResp.workstate;
    DEBUGLOG2("%010d-ComlinkR_TxCommandEx: BEFIPR response received, dataLen=%d, Status=%d", TO_UDINT(rc-4), pStatus^$UDINT);
    //DEBUG_VERBOSE3("%010d-                    uiLng=%d, aData[0]=0x%08X, aData[4]=0x%08X", TO_UDINT(pLogin^.befiprResp.resu.uiLng), pLogin^.befiprResp.resu.aData[0]$UDINT, pLogin^.befiprResp.resu.aData[4]$UDINT);
    retval := COMLINK_IPR;
  END_IF;

END_FUNCTION

//------------------------------------------------------------------------------
// ComlinkR_TxUpd_nocs
//------------------------------------------------------------------------------
FUNCTION ComlinkR_TxUpd_nocs
VAR_INPUT
    pLslcommregdata : ^lslCommregData;
    pLogin          : ^loginContextR; // connection context
    uiflags         : UINT;
END_VAR
VAR_OUTPUT
    retval          : comlinkReason;
END_VAR
VAR
    pt_comStCell  : ^comStCell;
    updList       : ^updateList;
    listIndex     : UDINT;
    listType      : UDINT;
    reqMsg        : msgTxUpdReqData;   // request structure for command CMD_TXUPD
    timx           : udint;
END_VAR

  retval := COMLINK_ERR_GENERAL;

  IF pLslcommregdata^.varpos$INT < 1000 THEN
    updList   := #pLogin^.statList;
    listIndex := pLslcommregdata^.varpos;
    listType  := 0;
  ELSE
    updList   := #pLogin^.dynList;
    listIndex := pLslcommregdata^.varpos - 1000;
    listType  := 1;
  END_IF;

  IF listIndex >= updList^.nbrCells THEN
    IF IncreaseUpdateList(updList, listIndex + 1, listType) = NIL THEN
      DEBUGLOG0("%010d-*** ComlinkR_TxUpd: MemoryUpdateList failed");
      DisconnectAfterErrorR(pLogin);
      RETURN;
    END_IF;
    DEBUGLOG2("%010d-*** ComlinkR_TxUpd: list %d increased to %d entries", listType, updList^.nbrCells);
  END_IF;

  pt_comStCell := updList^.pFirstCell + (listIndex * SIZEOF (comStCell));

  timx                       := pLslcommregdata^.uiTime; // u32 := u16
  pt_comStCell^.dData        := 16#80000001$DINT;     // INVALID
  pt_comStCell^.pCh          := pLslcommregdata^.LASALID$^SVRCH;
  pt_comStCell^.udUpdateRate := (timx and 16#3FFF) or ((timx and 16#C000) shl 16) or (uiflags shl 14);
  pt_comStCell^.VarlistID    := pLslcommregdata^.VarlistID;
  pt_comStCell^.udLastUpdate := 0;

  reqMsg.iOff    := pLslcommregdata^.varpos$UINT;
  reqMsg.comcell := pt_comStCell^;  // copy struct on struct;
  // Send the request
  retval := SendRequestR(pLogin,
                         CMD_TXUPD,
                         respRequired:=FALSE,
                         #reqMsg,
                         SIZEOF(reqMsg),
                         blockingMode:=TRUE);
  IF retval = 0 THEN
    DEBUGLOG1("%010d-    ComlinkR_TxUpd_nocs: sent cell ofs %d", TO_UDINT(reqMsg.iOff));
  ELSE
    DEBUGLOG1("%010d-*** ComlinkR_TxUpd_nocs: SendRequestR failed, retval=%d", TO_UDINT(retval));
  END_IF;

END_FUNCTION

//------------------------------------------------------------------------------
// ComlinkR_TxUpd
//
// Return value:
//  If the function succeeds, the return value is 0, othzerwise it is a
//  negative error code.
//------------------------------------------------------------------------------
FUNCTION ComlinkR_TxUpd
VAR_INPUT
    pLslcommregdata : ^lslCommregData;
    pComdef         : ^comdef;
    res             : UDINT;
    uiflags         : UINT;
END_VAR
VAR_OUTPUT
    retval          : comlinkReason;
END_VAR
VAR
    pLogin          : ^loginContextR; // connection context
END_VAR

  IF !!isComlinkRInitialized THEN
    retval := COMLINK_ERR_CLIENT_NOTREADY;
    RETURN;
  END_IF;

  pLogin := pComdef^$comdefT.pLogin$^loginContextR;
  IF pLogin = NIL THEN
    retval := COMLINK_ERR_LOGIN_REQUIRED;
    RETURN;
  END_IF;

  retval := ComlinkR_TxUpd_nocs(pLslcommregdata, pLogin, uiflags);

END_FUNCTION

//------------------------------------------------------------------------------
// SendMaxIdleTime_RS232_nocs
//------------------------------------------------------------------------------
FUNCTION SendMaxIdleTime_RS232_nocs
VAR_INPUT
  pComdefT : ^comdefT;
  remoteMaxIdleTime_ms : UDINT;
  pLogin          : ^loginContextR; // connection context
END_VAR
VAR_OUTPUT
  retVal : DINT;
END_VAR
VAR
    reqMsg        : msgIdlTimReqData;  // request structure for command CMD_MAXIDLETIME
END_VAR

  //retval := COMLINK_ERR_GENERAL;

  // prepare the request message structure
  reqMsg.maxIdleTime_ms := remoteMaxIdleTime_ms;

  // Send the request
  retval := SendRequestR(pLogin,
                         CMD_MAXIDLETIME,
                         respRequired:=FALSE,
                         #reqMsg,
                         SIZEOF(reqMsg),
                         blockingMode:=TRUE);
  IF retval = 0 THEN
    DEBUGLOG0("%010d-SendMaxIdleTime_RS232_nocs: MAXIDLETIME request sent");
  ELSE
    DEBUGLOG1("%010d-*** SendMaxIdleTime_RS232_nocs: SendCmdMsg failed, rc=%d", TO_UDINT(retval));
  END_IF;

END_FUNCTION

//------------------------------------------------------------------------------
// SendMaxIdleTime_RS232
//
// Return value:
//  If the function succeeds, the return value is 0, othzerwise it is a
//  negative error code.
//------------------------------------------------------------------------------
FUNCTION SendMaxIdleTime_RS232
VAR_INPUT
  pComdefT : ^comdefT;
  remoteMaxIdleTime_ms : UDINT;
END_VAR
VAR_OUTPUT
  retVal : DINT;
END_VAR
VAR
    pLogin          : ^loginContextR; // connection context
END_VAR

  IF !!isComlinkRInitialized THEN
    retval := COMLINK_ERR_CLIENT_NOTREADY;
    RETURN;
  END_IF;

  pLogin := pComdefT^.pLogin$^loginContextR;
  IF pLogin = NIL THEN
    retval := COMLINK_ERR_LOGIN_REQUIRED;
    RETURN;
  END_IF;

  retval := SendMaxIdleTime_RS232_nocs(pComdefT, remoteMaxIdleTime_ms, pLogin);

END_FUNCTION

//------------------------------------------------------------------------------
// ComlinkR_InstallCallback
//------------------------------------------------------------------------------
FUNCTION ComlinkR_InstallCallback
VAR_INPUT
    pCallback : ^void;
END_VAR
VAR
    i         : UDINT;
    pLogin    : ^loginContextR;
END_VAR

  IF !!isComlinkRInitialized THEN
    RETURN;
  END_IF;

  DEBUGLOG1("%010d-ComlinkR_InstallCallback: pCallback=0x%08X", pCallback$UDINT);

  FOR i := 0 TO (arraysize(loginArrayR) - 1) DO
    pLogin := loginArrayR[i];
    IF pLogin <> NIL & pLogin^.isClient THEN
      pLogin^.pCallback := pCallback;
    END_IF;
  END_FOR;

  g_pCallback := pCallback;

END_FUNCTION

//------------------------------------------------------------------------------
// ComlinkR_StartStopRefresh_nocs
//------------------------------------------------------------------------------
FUNCTION ComlinkR_StartStopRefresh_nocs
VAR_INPUT
    pLogin   : ^loginContextR; // connection context
    count    : UINT;
    typ      : UINT;
    res      : UDINT;
END_VAR
VAR_OUTPUT
    retval    : comlinkReason;
END_VAR
VAR
    reqMsg        : msgSsRefrReqData;  // request structure for command CMD_SSREFR
END_VAR

//  retval := COMLINK_ERR_GENERAL;

  // prepare the request message structure
  reqMsg.count   := count;
  reqMsg.typ     := typ;

  // Send the request
  retval := SendRequestR(pLogin,
                         CMD_SSREFR,
                         respRequired:=FALSE,
                         #reqMsg,
                         SIZEOF(reqMsg),
                         blockingMode:=TRUE);
  IF retval = 0 THEN
    DEBUGLOG3("%010d-ComlinkR_StartStopRefresh: SSREFR request sent, msgLen=%d, typ=%d, count=%d", TO_UDINT(retval), TO_UDINT(typ), TO_UDINT(count));
  ELSE
    DEBUGLOG3("%010d-*** ComlinkR_StartStopRefresh(typ %d, count %d): SendRequestR failed, rc=%d", TO_UDINT(typ), TO_UDINT(count), TO_UDINT(retval));
  END_IF;

END_FUNCTION

//------------------------------------------------------------------------------
// ComlinkR_StartStopRefresh
//------------------------------------------------------------------------------
FUNCTION ComlinkR_StartStopRefresh
VAR_INPUT
    pComdef  : ^comdef;
    count    : UINT;
    typ      : UINT;
    res      : UDINT;
END_VAR
VAR_OUTPUT
    retval   : comlinkReason;
END_VAR
VAR
    pLogin        : ^loginContextR; // connection context
END_VAR

  IF !!isComlinkRInitialized THEN
    retval := COMLINK_ERR_CLIENT_NOTREADY;
    RETURN;
  END_IF;

  pLogin := pComdef^$comdefT.pLogin$^loginContextR;
  IF pLogin = NIL THEN
    retval := COMLINK_ERR_LOGIN_REQUIRED;
    RETURN;
  END_IF;

  retval := ComlinkR_StartStopRefresh_nocs(pLogin, count, typ, res);

END_FUNCTION

//------------------------------------------------------------------------------
// UpdateCell
//
// Return value:
//  Error                                                     : <=0
//  When udLastUpdate did not expire                          : 1
//  When udLastUpdate expired, but dData did not change       : 2
//  When udLastUpdate expired, and dData changed (transfer)   : 3
//------------------------------------------------------------------------------
FUNCTION UpdateCellR
VAR_INPUT
    pLogin : ^loginContextR;
    pUpdCell      : ^comStCell;  // pointer to cell in updatelist
    iOff          : UINT;
END_VAR
VAR_OUTPUT
    retval        : DINT;
END_VAR
VAR
    reqMsg        : msgUpdCellReqData; // request structure for command CMD_UPDCELL
    dData         : DINT;
    rc            : UINT;
END_VAR
